    CONST robtarget Target_LetFron3_660:=[[-82.267,-107.387,45.753],[0.430645927,0.216920311,0.57802214,0.658316087],[0,0,0,0],[9E+09,9E+09,9E+09,9E+09,9E+09,9E+09]];
    CONST robtarget Target_LetFron3_670:=[[-81.504,-107.822,44.831],[0.430645927,0.216920311,0.57802214,0.658316087],[0,0,0,0],[9E+09,9E+09,9E+09,9E+09,9E+09,9E+09]];
    CONST robtarget Target_LetFron3_680:=[[-81.6,-107.767,55.109],[0.430645927,0.216920311,0.57802214,0.658316087],[0,0,0,0],[9E+09,9E+09,9E+09,9E+09,9E+09,9E+09]];
    CONST robtarget Target_LetFron3_690:=[[-91.637,-127.746,55.109],[0.430645927,0.216920311,0.57802214,0.658316087],[0,0,0,0],[9E+09,9E+09,9E+09,9E+09,9E+09,9E+09]];
    CONST robtarget Target_LetFron3_700:=[[-88.514,-129.459,54.672],[0.430645927,0.216920311,0.57802214,0.658316087],[0,0,0,0],[9E+09,9E+09,9E+09,9E+09,9E+09,9E+09]];
    CONST robtarget Target_LetFron3_710:=[[-78.514,-109.459,54.672],[0.430645927,0.216920311,0.57802214,0.658316087],[0,0,0,0],[9E+09,9E+09,9E+09,9E+09,9E+09,9E+09]];
    CONST robtarget Target_LetFron3_720:=[[-77.118,-110.187,55.177],[0.430645927,0.216920311,0.57802214,0.658316087],[0,0,0,0],[9E+09,9E+09,9E+09,9E+09,9E+09,9E+09]];
    CONST robtarget Target_LetFron3_730:=[[-75.152,-111.175,55.401],[0.430645927,0.216920311,0.57802214,0.658316087],[0,0,0,0],[9E+09,9E+09,9E+09,9E+09,9E+09,9E+09]];
    CONST robtarget Target_LetFron3_740:=[[-73.482,-111.981,54.982],[0.430645927,0.216920311,0.57802214,0.658316087],[0,0,0,0],[9E+09,9E+09,9E+09,9E+09,9E+09,9E+09]];
    CONST robtarget Target_LetFron3_750:=[[-72.199,-112.579,54.044],[0.430645927,0.216920311,0.57802214,0.658316087],[0,0,0,0],[9E+09,9E+09,9E+09,9E+09,9E+09,9E+09]];
    CONST robtarget Target_LetFron3_760:=[[-71.586,-112.859,52.943],[0.430645927,0.216920311,0.57802214,0.658316087],[0,0,0,0],[9E+09,9E+09,9E+09,9E+09,9E+09,9E+09]];
    CONST robtarget Target_LetFron3_770:=[[-71.209,-113.029,51.815],[0.430645927,0.216920311,0.57802214,0.658316087],[0,0,0,0],[9E+09,9E+09,9E+09,9E+09,9E+09,9E+09]];
    CONST robtarget Target_LetFron3_780:=[[-71.14,-113.06,50.668],[0.430645927,0.216920311,0.57802214,0.658316087],[0,0,0,0],[9E+09,9E+09,9E+09,9E+09,9E+09,9E+09]];
    CONST robtarget Target_LetFron3_790:=[[-71.14,-113.06,49.432],[0.430645927,0.216920311,0.57802214,0.658316087],[0,0,0,0],[9E+09,9E+09,9E+09,9E+09,9E+09,9E+09]];
    CONST robtarget Target_LetFron3_800:=[[-71.288,-112.994,48.254],[0.430645927,0.216920311,0.57802214,0.658316087],[0,0,0,0],[9E+09,9E+09,9E+09,9E+09,9E+09,9E+09]];
    CONST robtarget Target_LetFron3_810:=[[-71.728,-112.794,47.133],[0.430645927,0.216920311,0.57802214,0.658316087],[0,0,0,0],[9E+09,9E+09,9E+09,9E+09,9E+09,9E+09]];
    CONST robtarget Target_LetFron3_820:=[[-72.376,-112.498,46.001],[0.430645927,0.216920311,0.57802214,0.658316087],[0,0,0,0],[9E+09,9E+09,9E+09,9E+09,9E+09,9E+09]];
    CONST robtarget Target_LetFron3_830:=[[-73.318,-112.058,45.279],[0.430645927,0.216920311,0.57802214,0.658316087],[0,0,0,0],[9E+09,9E+09,9E+09,9E+09,9E+09,9E+09]];
    CONST robtarget Target_LetFron3_840:=[[-74.681,-111.405,44.719],[0.430645927,0.216920311,0.57802214,0.658316087],[0,0,0,0],[9E+09,9E+09,9E+09,9E+09,9E+09,9E+09]];
    CONST robtarget Target_LetFron3_850:=[[-75.902,-110.803,44.719],[0.430645927,0.216920311,0.57802214,0.658316087],[0,0,0,0],[9E+09,9E+09,9E+09,9E+09,9E+09,9E+09]];
    CONST robtarget Target_LetFron3_860:=[[-77.054,-110.22,45.141],[0.430645927,0.216920311,0.57802214,0.658316087],[0,0,0,0],[9E+09,9E+09,9E+09,9E+09,9E+09,9E+09]];
    CONST robtarget Target_LetFron3_870:=[[-77.919,-109.772,46.005],[0.430645927,0.216920311,0.57802214,0.658316087],[0,0,0,0],[9E+09,9E+09,9E+09,9E+09,9E+09,9E+09]];
    CONST robtarget Target_LetFron3_880:=[[-78.398,-109.52,46.991],[0.430645927,0.216920311,0.57802214,0.658316087],[0,0,0,0],[9E+09,9E+09,9E+09,9E+09,9E+09,9E+09]];
    CONST robtarget Target_LetFron3_890:=[[-78.609,-109.408,48.208],[0.430645927,0.216920311,0.57802214,0.658316087],[0,0,0,0],[9E+09,9E+09,9E+09,9E+09,9E+09,9E+09]];
    CONST robtarget Target_LetFron3_900:=[[-78.594,-109.416,49.608],[0.430645927,0.216920311,0.57802214,0.658316087],[0,0,0,0],[9E+09,9E+09,9E+09,9E+09,9E+09,9E+09]];
    CONST robtarget Target_LetFron3_910:=[[-78.574,-109.427,49.862],[0.430645927,0.216920311,0.57802214,0.658316087],[0,0,0,0],[9E+09,9E+09,9E+09,9E+09,9E+09,9E+09]];
    CONST robtarget Target_LetFron3_920:=[[-77.106,-110.19,49.869],[0.430645927,0.216920311,0.57802214,0.658316087],[0,0,0,0],[9E+09,9E+09,9E+09,9E+09,9E+09,9E+09]];
    CONST robtarget Target_LetFron3_930:=[[-72.898,-112.255,49.869],[0.430645927,0.216920311,0.57802214,0.658316087],[0,0,0,0],[9E+09,9E+09,9E+09,9E+09,9E+09,9E+09]];
    CONST robtarget Target_LetFron3_940:=[[-82.898,-132.255,49.869],[0.430645927,0.216920311,0.57802214,0.658316087],[0,0,0,0],[9E+09,9E+09,9E+09,9E+09,9E+09,9E+09]];
    CONST robtarget Target_LetFron3_950:=[[-80.313,-133.427,54.778],[0.430645927,0.216920311,0.57802214,0.658316087],[0,0,0,0],[9E+09,9E+09,9E+09,9E+09,9E+09,9E+09]];
    CONST robtarget Target_LetFron3_960:=[[-70.313,-113.427,54.778],[0.430645927,0.216920311,0.57802214,0.658316087],[0,0,0,0],[9E+09,9E+09,9E+09,9E+09,9E+09,9E+09]];
    CONST robtarget Target_LetFron3_970:=[[-68.992,-113.999,55.279],[0.430645927,0.216920311,0.57802214,0.658316087],[0,0,0,0],[9E+09,9E+09,9E+09,9E+09,9E+09,9E+09]];
    CONST robtarget Target_LetFron3_980:=[[-67.664,-114.556,55.401],[0.430645927,0.216920311,0.57802214,0.658316087],[0,0,0,0],[9E+09,9E+09,9E+09,9E+09,9E+09,9E+09]];
    CONST robtarget Target_LetFron3_990:=[[-66.498,-115.03,55.08],[0.430645927,0.216920311,0.57802214,0.658316087],[0,0,0,0],[9E+09,9E+09,9E+09,9E+09,9E+09,9E+09]];
    CONST robtarget Target_LetFron3_1000:=[[-65.468,-115.437,54.06],[0.430645927,0.216920311,0.57802214,0.658316087],[0,0,0,0],[9E+09,9E+09,9E+09,9E+09,9E+09,9E+09]];
    CONST robtarget Target_LetFron3_1010:=[[-65.245,-115.524,53.314],[0.430645927,0.216920311,0.57802214,0.658316087],[0,0,0,0],[9E+09,9E+09,9E+09,9E+09,9E+09,9E+09]];
    CONST robtarget Target_LetFron3_1020:=[[-65.368,-115.476,43.276],[0.430645927,0.216920311,0.57802214,0.658316087],[0,0,0,0],[9E+09,9E+09,9E+09,9E+09,9E+09,9E+09]];
    CONST robtarget Target_LetFron3_1030:=[[-65.313,-115.498,44.991],[0.430645927,0.216920311,0.57802214,0.658316087],[0,0,0,0],[9E+09,9E+09,9E+09,9E+09,9E+09,9E+09]];
    CONST robtarget Target_LetFron3_1040:=[[-63.93,-116.026,45.188],[0.430645927,0.216920311,0.57802214,0.658316087],[0,0,0,0],[9E+09,9E+09,9E+09,9E+09,9E+09,9E+09]];
    CONST robtarget Target_LetFron3_1050:=[[-70.13,-113.508,44.989],[0.430645927,0.216920311,0.57802214,0.658316087],[0,0,0,0],[9E+09,9E+09,9E+09,9E+09,9E+09,9E+09]];
    CONST robtarget Target_LetFron3_1060:=[[-80.13,-133.508,44.989],[0.430645927,0.216920311,0.57802214,0.658316087],[0,0,0,0],[9E+09,9E+09,9E+09,9E+09,9E+09,9E+09]];
    CONST robtarget Target_LetFron3_1070:=[[-72.339,-136.611,45.952],[0.430645927,0.216920311,0.57802214,0.658316087],[0,0,0,0],[9E+09,9E+09,9E+09,9E+09,9E+09,9E+09]];
    CONST robtarget Target_LetFron3_1080:=[[-62.36,-116.604,45.863],[0.430645927,0.216920311,0.57802214,0.658316087],[0,0,0,0],[9E+09,9E+09,9E+09,9E+09,9E+09,9E+09]];
    CONST robtarget Target_LetFron3_1090:=[[-60.366,-117.303,44.736],[0.430645927,0.216920311,0.57802214,0.658316087],[0,0,0,0],[9E+09,9E+09,9E+09,9E+09,9E+09,9E+09]];
    CONST robtarget Target_LetFron3_1100:=[[-58.61,-117.888,44.82],[0.430645927,0.216920311,0.57802214,0.658316087],[0,0,0,0],[9E+09,9E+09,9E+09,9E+09,9E+09,9E+09]];
    CONST robtarget Target_LetFron3_1110:=[[-56.667,-118.501,45.956],[0.430645927,0.216920311,0.57802214,0.658316087],[0,0,0,0],[9E+09,9E+09,9E+09,9E+09,9E+09,9E+09]];
    CONST robtarget Target_LetFron3_1120:=[[-56.029,-118.695,47.133],[0.430645927,0.216920311,0.57802214,0.658316087],[0,0,0,0],[9E+09,9E+09,9E+09,9E+09,9E+09,9E+09]];
    CONST robtarget Target_LetFron3_1130:=[[-56.121,-118.667,48.621],[0.430645927,0.216920311,0.57802214,0.658316087],[0,0,0,0],[9E+09,9E+09,9E+09,9E+09,9E+09,9E+09]];
    CONST robtarget Target_LetFron3_1140:=[[-56.545,-118.539,49.359],[0.430645927,0.216920311,0.57802214,0.658316087],[0,0,0,0],[9E+09,9E+09,9E+09,9E+09,9E+09,9E+09]];
    CONST robtarget Target_LetFron3_1150:=[[-57.437,-118.262,50.034],[0.430645927,0.216920311,0.57802214,0.658316087],[0,0,0,0],[9E+09,9E+09,9E+09,9E+09,9E+09,9E+09]];
    CONST robtarget Target_LetFron3_1160:=[[-58.505,-117.922,50.535],[0.430645927,0.216920311,0.57802214,0.658316087],[0,0,0,0],[9E+09,9E+09,9E+09,9E+09,9E+09,9E+09]];
    CONST robtarget Target_LetFron3_1170:=[[-59.869,-117.471,51.117],[0.430645927,0.216920311,0.57802214,0.658316087],[0,0,0,0],[9E+09,9E+09,9E+09,9E+09,9E+09,9E+09]];
    CONST robtarget Target_LetFron3_1180:=[[-60.318,-117.319,51.376],[0.430645927,0.216920311,0.57802214,0.658316087],[0,0,0,0],[9E+09,9E+09,9E+09,9E+09,9E+09,9E+09]];
    CONST robtarget Target_LetFron3_1190:=[[-62.669,-116.492,52.048],[0.430645927,0.216920311,0.57802214,0.658316087],[0,0,0,0],[9E+09,9E+09,9E+09,9E+09,9E+09,9E+09]];
    CONST robtarget Target_LetFron3_1200:=[[-62.602,-116.516,52.834],[0.430645927,0.216920311,0.57802214,0.658316087],[0,0,0,0],[9E+09,9E+09,9E+09,9E+09,9E+09,9E+09]];
    CONST robtarget Target_LetFron3_1210:=[[-62.228,-116.651,53.814],[0.430645927,0.216920311,0.57802214,0.658316087],[0,0,0,0],[9E+09,9E+09,9E+09,9E+09,9E+09,9E+09]];
    CONST robtarget Target_LetFron3_1220:=[[-61.449,-116.928,54.619],[0.430645927,0.216920311,0.57802214,0.658316087],[0,0,0,0],[9E+09,9E+09,9E+09,9E+09,9E+09,9E+09]];
    CONST robtarget Target_LetFron3_1230:=[[-60.216,-117.353,55.205],[0.430645927,0.216920311,0.57802214,0.658316087],[0,0,0,0],[9E+09,9E+09,9E+09,9E+09,9E+09,9E+09]];
    CONST robtarget Target_LetFron3_1240:=[[-58.271,-117.997,55.4],[0.430645927,0.216920311,0.57802214,0.658316087],[0,0,0,0],[9E+09,9E+09,9E+09,9E+09,9E+09,9E+09]];
    CONST robtarget Target_LetFron3_1250:=[[-56.602,-118.521,55.079],[0.430645927,0.216920311,0.57802214,0.658316087],[0,0,0,0],[9E+09,9E+09,9E+09,9E+09,9E+09,9E+09]];
    CONST robtarget Target_LetFron3_1260:=[[-55.798,-118.764,54.785],[0.430645927,0.216920311,0.57802214,0.658316087],[0,0,0,0],[9E+09,9E+09,9E+09,9E+09,9E+09,9E+09]];
    CONST robtarget Target_LetFron3_1270:=[[-65.797,-138.765,54.792],[0.430645927,0.216920311,0.57802214,0.658316087],[0,0,0,0],[9E+09,9E+09,9E+09,9E+09,9E+09,9E+09]];
    CONST robtarget Target_LetFron3_1280:=[[-62.847,-139.607,55.109],[0.430645927,0.216920311,0.57802214,0.658316087],[0,0,0,0],[9E+09,9E+09,9E+09,9E+09,9E+09,9E+09]];
    CONST robtarget Target_LetFron3_1290:=[[-52.847,-119.607,55.109],[0.430645927,0.216920311,0.57802214,0.658316087],[0,0,0,0],[9E+09,9E+09,9E+09,9E+09,9E+09,9E+09]];
    CONST robtarget Target_LetFron3_1300:=[[-52.608,-119.672,44.874],[0.430645927,0.216920311,0.57802214,0.658316087],[0,0,0,0],[9E+09,9E+09,9E+09,9E+09,9E+09,9E+09]];
    CONST robtarget Target_LetFron3_1310:=[[-62.608,-139.672,44.874],[0.430645927,0.216920311,0.57802214,0.658316087],[0,0,0,0],[9E+09,9E+09,9E+09,9E+09,9E+09,9E+09]];
    CONST robtarget Target_LetFron3_1320:=[[-62.417,-139.723,40.356],[0.430645927,0.216920311,0.57802214,0.658316087],[0,0,0,0],[9E+09,9E+09,9E+09,9E+09,9E+09,9E+09]];
    CONST robtarget Target_LetFron3_1330:=[[-52.574,-119.681,40.311],[0.430645927,0.216920311,0.57802214,0.658316087],[0,0,0,0],[9E+09,9E+09,9E+09,9E+09,9E+09,9E+09]];
    CONST robtarget Target_LetFron3_1340:=[[-62.574,-139.681,40.311],[0.430645927,0.216920311,0.57802214,0.658316087],[0,0,0,0],[9E+09,9E+09,9E+09,9E+09,9E+09,9E+09]];
    CONST robtarget Target_LetFron3_1350:=[[-58.595,-140.685,42.493],[0.430645927,0.216920311,0.57802214,0.658316087],[0,0,0,0],[9E+09,9E+09,9E+09,9E+09,9E+09,9E+09]];
    CONST robtarget Target_LetFron3_1360:=[[-48.595,-120.685,42.493],[0.430645927,0.216920311,0.57802214,0.658316087],[0,0,0,0],[9E+09,9E+09,9E+09,9E+09,9E+09,9E+09]];
    CONST robtarget Target_LetFron3_1370:=[[-42.535,-121.952,41.813],[0.430645927,0.216920311,0.57802214,0.658316087],[0,0,0,0],[9E+09,9E+09,9E+09,9E+09,9E+09,9E+09]];
    CONST robtarget Target_LetFron3_1380:=[[-41.416,-122.152,42.942],[0.430645927,0.216920311,0.57802214,0.658316087],[0,0,0,0],[9E+09,9E+09,9E+09,9E+09,9E+09,9E+09]];
    CONST robtarget Target_LetFron3_1390:=[[-40.861,-122.247,44.157],[0.430645927,0.216920311,0.57802214,0.658316087],[0,0,0,0],[9E+09,9E+09,9E+09,9E+09,9E+09,9E+09]];
    CONST robtarget Target_LetFron3_1400:=[[-40.861,-122.247,45.481],[0.430645927,0.216920311,0.57802214,0.658316087],[0,0,0,0],[9E+09,9E+09,9E+09,9E+09,9E+09,9E+09]];
    CONST robtarget Target_LetFron3_1410:=[[-41.204,-122.188,46.641],[0.430645927,0.216920311,0.57802214,0.658316087],[0,0,0,0],[9E+09,9E+09,9E+09,9E+09,9E+09,9E+09]];
    CONST robtarget Target_LetFron3_1420:=[[-41.998,-122.049,47.583],[0.430645927,0.216920311,0.57802214,0.658316087],[0,0,0,0],[9E+09,9E+09,9E+09,9E+09,9E+09,9E+09]];
    CONST robtarget Target_LetFron3_1430:=[[-43.35,-121.797,48.403],[0.430645927,0.216920311,0.57802214,0.658316087],[0,0,0,0],[9E+09,9E+09,9E+09,9E+09,9E+09,9E+09]];
    CONST robtarget Target_LetFron3_1440:=[[-44.844,-121.506,49.112],[0.430645927,0.216920311,0.57802214,0.658316087],[0,0,0,0],[9E+09,9E+09,9E+09,9E+09,9E+09,9E+09]];
    CONST robtarget Target_LetFron3_1450:=[[-46.229,-121.217,49.939],[0.430645927,0.216920311,0.57802214,0.658316087],[0,0,0,0],[9E+09,9E+09,9E+09,9E+09,9E+09,9E+09]];
    CONST robtarget Target_LetFron3_1460:=[[-49.035,-120.581,50.611],[0.430645927,0.216920311,0.57802214,0.658316087],[0,0,0,0],[9E+09,9E+09,9E+09,9E+09,9E+09,9E+09]];
    CONST robtarget Target_LetFron3_1470:=[[-48.955,-120.6,52.318],[0.430645927,0.216920311,0.57802214,0.658316087],[0,0,0,0],[9E+09,9E+09,9E+09,9E+09,9E+09,9E+09]];
    CONST robtarget Target_LetFron3_1480:=[[-48.452,-120.719,53.355],[0.430645927,0.216920311,0.57802214,0.658316087],[0,0,0,0],[9E+09,9E+09,9E+09,9E+09,9E+09,9E+09]];
    CONST robtarget Target_LetFron3_1490:=[[-47.435,-120.951,54.415],[0.430645927,0.216920311,0.57802214,0.658316087],[0,0,0,0],[9E+09,9E+09,9E+09,9E+09,9E+09,9E+09]];
    CONST robtarget Target_LetFron3_1500:=[[-45.861,-121.294,55.128],[0.430645927,0.216920311,0.57802214,0.658316087],[0,0,0,0],[9E+09,9E+09,9E+09,9E+09,9E+09,9E+09]];
    CONST robtarget Target_LetFron3_1510:=[[-43.532,-121.765,55.401],[0.430645927,0.216920311,0.57802214,0.658316087],[0,0,0,0],[9E+09,9E+09,9E+09,9E+09,9E+09,9E+09]];
    CONST robtarget Target_LetFron3_1520:=[[-41.726,-122.098,55.154],[0.430645927,0.216920311,0.57802214,0.658316087],[0,0,0,0],[9E+09,9E+09,9E+09,9E+09,9E+09,9E+09]];
    CONST robtarget Target_LetFron3_1530:=[[-40.575,-122.295,54.72],[0.430645927,0.216920311,0.57802214,0.658316087],[0,0,0,0],[9E+09,9E+09,9E+09,9E+09,9E+09,9E+09]];
    CONST robtarget Target_LetFron3_1540:=[[-50.576,-142.295,54.717],[0.430645927,0.216920311,0.57802214,0.658316087],[0,0,0,0],[9E+09,9E+09,9E+09,9E+09,9E+09,9E+09]];
    CONST robtarget Target_LetFron3_1550:=[[-43.98,-143.216,54.592],[0.430645927,0.216920311,0.57802214,0.658316087],[0,0,0,0],[9E+09,9E+09,9E+09,9E+09,9E+09,9E+09]];
    CONST robtarget Target_LetFron3_1560:=[[-33.98,-123.216,54.592],[0.430645927,0.216920311,0.57802214,0.658316087],[0,0,0,0],[9E+09,9E+09,9E+09,9E+09,9E+09,9E+09]];
    CONST robtarget Target_LetFron3_1570:=[[-32.448,-123.378,55.116],[0.430645927,0.216920311,0.57802214,0.658316087],[0,0,0,0],[9E+09,9E+09,9E+09,9E+09,9E+09,9E+09]];
    CONST robtarget Target_LetFron3_1580:=[[-30.55,-123.554,55.401],[0.430645927,0.216920311,0.57802214,0.658316087],[0,0,0,0],[9E+09,9E+09,9E+09,9E+09,9E+09,9E+09]];
    CONST robtarget Target_LetFron3_1590:=[[-28.936,-123.68,55.282],[0.430645927,0.216920311,0.57802214,0.658316087],[0,0,0,0],[9E+09,9E+09,9E+09,9E+09,9E+09,9E+09]];
    CONST robtarget Target_LetFron3_1600:=[[-27.719,-123.761,54.742],[0.430645927,0.216920311,0.57802214,0.658316087],[0,0,0,0],[9E+09,9E+09,9E+09,9E+09,9E+09,9E+09]];
    CONST robtarget Target_LetFron3_1610:=[[-26.596,-123.826,53.8],[0.430645927,0.216920311,0.57802214,0.658316087],[0,0,0,0],[9E+09,9E+09,9E+09,9E+09,9E+09,9E+09]];
    CONST robtarget Target_LetFron3_1620:=[[-25.968,-123.857,52.688],[0.430645927,0.216920311,0.57802214,0.658316087],[0,0,0,0],[9E+09,9E+09,9E+09,9E+09,9E+09,9E+09]];
    CONST robtarget Target_LetFron3_1630:=[[-25.618,-123.874,50.949],[0.430645927,0.216920311,0.57802214,0.658316087],[0,0,0,0],[9E+09,9E+09,9E+09,9E+09,9E+09,9E+09]];
    CONST robtarget Target_LetFron3_1640:=[[-25.618,-123.874,49.368],[0.430645927,0.216920311,0.57802214,0.658316087],[0,0,0,0],[9E+09,9E+09,9E+09,9E+09,9E+09,9E+09]];
    CONST robtarget Target_LetFron3_1650:=[[-25.967,-123.858,47.76],[0.430645927,0.216920311,0.57802214,0.658316087],[0,0,0,0],[9E+09,9E+09,9E+09,9E+09,9E+09,9E+09]];
    CONST robtarget Target_LetFron3_1660:=[[-26.976,-123.805,46.001],[0.430645927,0.216920311,0.57802214,0.658316087],[0,0,0,0],[9E+09,9E+09,9E+09,9E+09,9E+09,9E+09]];
    CONST robtarget Target_LetFron3_1670:=[[-28.333,-123.722,45.081],[0.430645927,0.216920311,0.57802214,0.658316087],[0,0,0,0],[9E+09,9E+09,9E+09,9E+09,9E+09,9E+09]];
    CONST robtarget Target_LetFron3_1680:=[[-29.666,-123.626,44.719],[0.430645927,0.216920311,0.57802214,0.658316087],[0,0,0,0],[9E+09,9E+09,9E+09,9E+09,9E+09,9E+09]];
    CONST robtarget Target_LetFron3_1690:=[[-30.876,-123.526,44.719],[0.430645927,0.216920311,0.57802214,0.658316087],[0,0,0,0],[9E+09,9E+09,9E+09,9E+09,9E+09,9E+09]];
    CONST robtarget Target_LetFron3_1700:=[[-32.317,-123.392,45.206],[0.430645927,0.216920311,0.57802214,0.658316087],[0,0,0,0],[9E+09,9E+09,9E+09,9E+09,9E+09,9E+09]];
    CONST robtarget Target_LetFron3_1710:=[[-32.996,-123.323,45.821],[0.430645927,0.216920311,0.57802214,0.658316087],[0,0,0,0],[9E+09,9E+09,9E+09,9E+09,9E+09,9E+09]];
    CONST robtarget Target_LetFron3_1720:=[[-33.54,-123.265,46.556],[0.430645927,0.216920311,0.57802214,0.658316087],[0,0,0,0],[9E+09,9E+09,9E+09,9E+09,9E+09,9E+09]];
    CONST robtarget Target_LetFron3_1730:=[[-33.887,-123.226,47.949],[0.430645927,0.216920311,0.57802214,0.658316087],[0,0,0,0],[9E+09,9E+09,9E+09,9E+09,9E+09,9E+09]];
    CONST robtarget Target_LetFron3_1740:=[[-33.912,-123.223,49.284],[0.430645927,0.216920311,0.57802214,0.658316087],[0,0,0,0],[9E+09,9E+09,9E+09,9E+09,9E+09,9E+09]];
    CONST robtarget Target_LetFron3_1750:=[[-33.868,-123.228,49.869],[0.430645927,0.216920311,0.57802214,0.658316087],[0,0,0,0],[9E+09,9E+09,9E+09,9E+09,9E+09,9E+09]];
    CONST robtarget Target_LetFron3_1760:=[[-27.55,-123.772,49.869],[0.430645927,0.216920311,0.57802214,0.658316087],[0,0,0,0],[9E+09,9E+09,9E+09,9E+09,9E+09,9E+09]];
    CONST robtarget Target_LetFron3_1770:=[[-37.55,-143.772,49.897],[0.430645927,0.216920311,0.57802214,0.658316087],[0,0,0,0],[9E+09,9E+09,9E+09,9E+09,9E+09,9E+09]];
    CONST robtarget Target_LetFron3_1780:=[[-31.259,-143.994,45.099],[0.430645927,0.216920311,0.57802214,0.658316087],[0,0,0,0],[9E+09,9E+09,9E+09,9E+09,9E+09,9E+09]];
    CONST robtarget Target_LetFron3_1790:=[[-21.259,-123.994,45.14],[0.430645927,0.216920311,0.57802214,0.658316087],[0,0,0,0],[9E+09,9E+09,9E+09,9E+09,9E+09,9E+09]];
    CONST robtarget Target_LetFron3_1800:=[[-19.408,-123.999,44.719],[0.430645927,0.216920311,0.57802214,0.658316087],[0,0,0,0],[9E+09,9E+09,9E+09,9E+09,9E+09,9E+09]];
    CONST robtarget Target_LetFron3_1810:=[[-17.893,-123.982,44.831],[0.430645927,0.216920311,0.57802214,0.658316087],[0,0,0,0],[9E+09,9E+09,9E+09,9E+09,9E+09,9E+09]];
    CONST robtarget Target_LetFron3_1820:=[[-16.252,-123.944,45.604],[0.430645927,0.216920311,0.57802214,0.658316087],[0,0,0,0],[9E+09,9E+09,9E+09,9E+09,9E+09,9E+09]];
    CONST robtarget Target_LetFron3_1830:=[[-15.038,-123.901,46.903],[0.430645927,0.216920311,0.57802214,0.658316087],[0,0,0,0],[9E+09,9E+09,9E+09,9E+09,9E+09,9E+09]];
    CONST robtarget Target_LetFron3_1840:=[[-14.306,-123.87,48.941],[0.430645927,0.216920311,0.57802214,0.658316087],[0,0,0,0],[9E+09,9E+09,9E+09,9E+09,9E+09,9E+09]];
    CONST robtarget Target_LetFron3_1850:=[[-14.248,-123.868,50.838],[0.430645927,0.216920311,0.57802214,0.658316087],[0,0,0,0],[9E+09,9E+09,9E+09,9E+09,9E+09,9E+09]];
    CONST robtarget Target_LetFron3_1860:=[[-14.656,-123.886,52.859],[0.430645927,0.216920311,0.57802214,0.658316087],[0,0,0,0],[9E+09,9E+09,9E+09,9E+09,9E+09,9E+09]];
    CONST robtarget Target_LetFron3_1870:=[[-15.358,-123.914,54.174],[0.430645927,0.216920311,0.57802214,0.658316087],[0,0,0,0],[9E+09,9E+09,9E+09,9E+09,9E+09,9E+09]];
    CONST robtarget Target_LetFron3_1880:=[[-16.312,-123.946,54.884],[0.430645927,0.216920311,0.57802214,0.658316087],[0,0,0,0],[9E+09,9E+09,9E+09,9E+09,9E+09,9E+09]];
    CONST robtarget Target_LetFron3_1890:=[[-17.794,-123.981,55.401],[0.430645927,0.216920311,0.57802214,0.658316087],[0,0,0,0],[9E+09,9E+09,9E+09,9E+09,9E+09,9E+09]];
    CONST robtarget Target_LetFron3_1900:=[[-18.988,-123.996,55.337],[0.430645927,0.216920311,0.57802214,0.658316087],[0,0,0,0],[9E+09,9E+09,9E+09,9E+09,9E+09,9E+09]];
    CONST robtarget Target_LetFron3_1910:=[[-20.839,-123.997,54.644],[0.430645927,0.216920311,0.57802214,0.658316087],[0,0,0,0],[9E+09,9E+09,9E+09,9E+09,9E+09,9E+09]];
    CONST robtarget Target_LetFron3_1920:=[[-21.239,-123.994,54.414],[0.430645927,0.216920311,0.57802214,0.658316087],[0,0,0,0],[9E+09,9E+09,9E+09,9E+09,9E+09,9E+09]];
    CONST robtarget Target_LetFron3_1930:=[[-22.525,-123.974,55.243],[0.430645927,0.216920311,0.57802214,0.658316087],[0,0,0,0],[9E+09,9E+09,9E+09,9E+09,9E+09,9E+09]];
    CONST robtarget Target_LetFron3_1940:=[[-22.191,-123.98,39.777],[0.430645927,0.216920311,0.57802214,0.658316087],[0,0,0,0],[9E+09,9E+09,9E+09,9E+09,9E+09,9E+09]];
    CONST robtarget Target_LetFron3_1950:=[[-32.321,-143.978,39.756],[0.430645927,0.216920311,0.57802214,0.658316087],[0,0,0,0],[9E+09,9E+09,9E+09,9E+09,9E+09,9E+09]];
    CONST robtarget Target_LetFron3_1960:=[[-12.321,-144.978,-58.244],[0.443836724,0.190106418,0.616719914,0.621711396],[0,0,0,0],[9E+09,9E+09,9E+09,9E+09,9E+09,9E+09]];
    !***********************************************************
    !Dibujo cuarto cuadrante de letrero frontal
    CONST robtarget Target_LetFron4_10:=[[-8.95,-145.995,82.097],[0.503297686,0.226891536,0.589713525,0.58944858],[0,0,0,0],[9E+09,9E+09,9E+09,9E+09,9E+09,9E+09]];
    CONST robtarget Target_LetFron4_20:=[[-18.95,-125.995,82.097],[0.503297686,0.226891536,0.589713525,0.58944858],[0,0,0,0],[9E+09,9E+09,9E+09,9E+09,9E+09,9E+09]];
    CONST robtarget Target_LetFron4_30:=[[-19.003,-125.994,68.333],[0.503297686,0.226891536,0.589713525,0.58944858],[0,0,0,0],[9E+09,9E+09,9E+09,9E+09,9E+09,9E+09]];
    CONST robtarget Target_LetFron4_40:=[[-23.592,-125.948,68.333],[0.503297686,0.226891536,0.589713525,0.58944858],[0,0,0,0],[9E+09,9E+09,9E+09,9E+09,9E+09,9E+09]];
    CONST robtarget Target_LetFron4_50:=[[-25.245,-125.89,69.103],[0.503297686,0.226891536,0.589713525,0.58944858],[0,0,0,0],[9E+09,9E+09,9E+09,9E+09,9E+09,9E+09]];
    CONST robtarget Target_LetFron4_60:=[[-26.403,-125.836,70.475],[0.503297686,0.226891536,0.589713525,0.58944858],[0,0,0,0],[9E+09,9E+09,9E+09,9E+09,9E+09,9E+09]];
    CONST robtarget Target_LetFron4_70:=[[-26.7,-125.82,71.985],[0.503297686,0.226891536,0.589713525,0.58944858],[0,0,0,0],[9E+09,9E+09,9E+09,9E+09,9E+09,9E+09]];
    CONST robtarget Target_LetFron4_80:=[[-26.314,-125.84,73.908],[0.503297686,0.226891536,0.589713525,0.58944858],[0,0,0,0],[9E+09,9E+09,9E+09,9E+09,9E+09,9E+09]];
    CONST robtarget Target_LetFron4_90:=[[-24.963,-125.901,75.447],[0.503297686,0.226891536,0.589713525,0.58944858],[0,0,0,0],[9E+09,9E+09,9E+09,9E+09,9E+09,9E+09]];
    CONST robtarget Target_LetFron4_100:=[[-21.051,-125.996,76.407],[0.503297686,0.226891536,0.589713525,0.58944858],[0,0,0,0],[9E+09,9E+09,9E+09,9E+09,9E+09,9E+09]];
    CONST robtarget Target_LetFron4_110:=[[-22.431,-125.976,76.317],[0.503297686,0.226891536,0.589713525,0.58944858],[0,0,0,0],[9E+09,9E+09,9E+09,9E+09,9E+09,9E+09]];
    CONST robtarget Target_LetFron4_120:=[[-26.29,-125.841,82.097],[0.503297686,0.226891536,0.589713525,0.58944858],[0,0,0,0],[9E+09,9E+09,9E+09,9E+09,9E+09,9E+09]];
    CONST robtarget Target_LetFron4_130:=[[-36.29,-145.841,82.097],[0.503297686,0.226891536,0.589713525,0.58944858],[0,0,0,0],[9E+09,9E+09,9E+09,9E+09,9E+09,9E+09]];
    CONST robtarget Target_LetFron4_140:=[[-42.667,-145.355,82.283],[0.503297686,0.226891536,0.589713525,0.58944858],[0,0,0,0],[9E+09,9E+09,9E+09,9E+09,9E+09,9E+09]];
    CONST robtarget Target_LetFron4_150:=[[-32.667,-125.355,82.283],[0.503297686,0.226891536,0.589713525,0.58944858],[0,0,0,0],[9E+09,9E+09,9E+09,9E+09,9E+09,9E+09]];
    CONST robtarget Target_LetFron4_160:=[[-34.857,-125.114,82.316],[0.503297686,0.226891536,0.589713525,0.58944858],[0,0,0,0],[9E+09,9E+09,9E+09,9E+09,9E+09,9E+09]];
    CONST robtarget Target_LetFron4_170:=[[-36.701,-124.879,81.437],[0.503297686,0.226891536,0.589713525,0.58944858],[0,0,0,0],[9E+09,9E+09,9E+09,9E+09,9E+09,9E+09]];
    CONST robtarget Target_LetFron4_180:=[[-37.577,-124.758,80.559],[0.503297686,0.226891536,0.589713525,0.58944858],[0,0,0,0],[9E+09,9E+09,9E+09,9E+09,9E+09,9E+09]];
    CONST robtarget Target_LetFron4_190:=[[-38.397,-124.639,78.755],[0.503297686,0.226891536,0.589713525,0.58944858],[0,0,0,0],[9E+09,9E+09,9E+09,9E+09,9E+09,9E+09]];
    CONST robtarget Target_LetFron4_200:=[[-38.556,-124.615,76.834],[0.503297686,0.226891536,0.589713525,0.58944858],[0,0,0,0],[9E+09,9E+09,9E+09,9E+09,9E+09,9E+09]];
    CONST robtarget Target_LetFron4_210:=[[-38.535,-124.618,75.633],[0.503297686,0.226891536,0.589713525,0.58944858],[0,0,0,0],[9E+09,9E+09,9E+09,9E+09,9E+09,9E+09]];
    CONST robtarget Target_LetFron4_220:=[[-38.089,-124.684,74.246],[0.503297686,0.226891536,0.589713525,0.58944858],[0,0,0,0],[9E+09,9E+09,9E+09,9E+09,9E+09,9E+09]];
    CONST robtarget Target_LetFron4_230:=[[-37.456,-124.775,73.108],[0.503297686,0.226891536,0.589713525,0.58944858],[0,0,0,0],[9E+09,9E+09,9E+09,9E+09,9E+09,9E+09]];
    CONST robtarget Target_LetFron4_240:=[[-36.441,-124.914,72.314],[0.503297686,0.226891536,0.589713525,0.58944858],[0,0,0,0],[9E+09,9E+09,9E+09,9E+09,9E+09,9E+09]];
    CONST robtarget Target_LetFron4_250:=[[-35.37,-125.051,71.858],[0.503297686,0.226891536,0.589713525,0.58944858],[0,0,0,0],[9E+09,9E+09,9E+09,9E+09,9E+09,9E+09]];
    CONST robtarget Target_LetFron4_260:=[[-33.892,-125.226,71.706],[0.503297686,0.226891536,0.589713525,0.58944858],[0,0,0,0],[9E+09,9E+09,9E+09,9E+09,9E+09,9E+09]];
    CONST robtarget Target_LetFron4_270:=[[-32.661,-125.357,71.87],[0.503297686,0.226891536,0.589713525,0.58944858],[0,0,0,0],[9E+09,9E+09,9E+09,9E+09,9E+09,9E+09]];
    CONST robtarget Target_LetFron4_280:=[[-31.413,-125.478,72.359],[0.503297686,0.226891536,0.589713525,0.58944858],[0,0,0,0],[9E+09,9E+09,9E+09,9E+09,9E+09,9E+09]];
    CONST robtarget Target_LetFron4_290:=[[-30.454,-125.562,73.003],[0.503297686,0.226891536,0.589713525,0.58944858],[0,0,0,0],[9E+09,9E+09,9E+09,9E+09,9E+09,9E+09]];
    CONST robtarget Target_LetFron4_300:=[[-29.503,-125.638,74.523],[0.503297686,0.226891536,0.589713525,0.58944858],[0,0,0,0],[9E+09,9E+09,9E+09,9E+09,9E+09,9E+09]];
    CONST robtarget Target_LetFron4_310:=[[-29.14,-125.665,75.942],[0.503297686,0.226891536,0.589713525,0.58944858],[0,0,0,0],[9E+09,9E+09,9E+09,9E+09,9E+09,9E+09]];
    CONST robtarget Target_LetFron4_320:=[[-29.014,-125.675,77.239],[0.503297686,0.226891536,0.589713525,0.58944858],[0,0,0,0],[9E+09,9E+09,9E+09,9E+09,9E+09,9E+09]];
    CONST robtarget Target_LetFron4_330:=[[-29.16,-125.664,78.757],[0.503297686,0.226891536,0.589713525,0.58944858],[0,0,0,0],[9E+09,9E+09,9E+09,9E+09,9E+09,9E+09]];
    CONST robtarget Target_LetFron4_340:=[[-29.598,-125.631,80.028],[0.503297686,0.226891536,0.589713525,0.58944858],[0,0,0,0],[9E+09,9E+09,9E+09,9E+09,9E+09,9E+09]];
    CONST robtarget Target_LetFron4_350:=[[-30.232,-125.58,80.936],[0.503297686,0.226891536,0.589713525,0.58944858],[0,0,0,0],[9E+09,9E+09,9E+09,9E+09,9E+09,9E+09]];
    CONST robtarget Target_LetFron4_360:=[[-31.211,-125.496,81.782],[0.503297686,0.226891536,0.589713525,0.58944858],[0,0,0,0],[9E+09,9E+09,9E+09,9E+09,9E+09,9E+09]];
    CONST robtarget Target_LetFron4_370:=[[-32.734,-125.348,82.291],[0.503297686,0.226891536,0.589713525,0.58944858],[0,0,0,0],[9E+09,9E+09,9E+09,9E+09,9E+09,9E+09]];
    CONST robtarget Target_LetFron4_380:=[[-42.734,-145.348,82.291],[0.503297686,0.226891536,0.589713525,0.58944858],[0,0,0,0],[9E+09,9E+09,9E+09,9E+09,9E+09,9E+09]];
    CONST robtarget Target_LetFron4_390:=[[-53.051,-143.856,72.591],[0.492892784,0.289203693,0.528592352,0.627700607],[0,0,0,0],[9E+09,9E+09,9E+09,9E+09,9E+09,9E+09]];
    CONST robtarget Target_LetFron4_400:=[[-43.051,-123.856,72.591],[0.492892784,0.289203693,0.528592352,0.627700607],[0,0,0,0],[9E+09,9E+09,9E+09,9E+09,9E+09,9E+09]];
    CONST robtarget Target_LetFron4_410:=[[-45.7,-123.329,71.706],[0.492892784,0.289203693,0.528592352,0.627700607],[0,0,0,0],[9E+09,9E+09,9E+09,9E+09,9E+09,9E+09]];
    CONST robtarget Target_LetFron4_420:=[[-46.898,-123.072,71.822],[0.492892784,0.289203693,0.528592352,0.627700607],[0,0,0,0],[9E+09,9E+09,9E+09,9E+09,9E+09,9E+09]];
    CONST robtarget Target_LetFron4_430:=[[-48.129,-122.794,72.468],[0.492892784,0.289203693,0.528592352,0.627700607],[0,0,0,0],[9E+09,9E+09,9E+09,9E+09,9E+09,9E+09]];
    CONST robtarget Target_LetFron4_440:=[[-49.172,-122.548,73.865],[0.492892784,0.289203693,0.528592352,0.627700607],[0,0,0,0],[9E+09,9E+09,9E+09,9E+09,9E+09,9E+09]];
    CONST robtarget Target_LetFron4_450:=[[-49.762,-122.405,76.003],[0.492892784,0.289203693,0.528592352,0.627700607],[0,0,0,0],[9E+09,9E+09,9E+09,9E+09,9E+09,9E+09]];
    CONST robtarget Target_LetFron4_460:=[[-49.705,-122.419,78.093],[0.492892784,0.289203693,0.528592352,0.627700607],[0,0,0,0],[9E+09,9E+09,9E+09,9E+09,9E+09,9E+09]];
    CONST robtarget Target_LetFron4_470:=[[-49.07,-122.573,80.012],[0.492892784,0.289203693,0.528592352,0.627700607],[0,0,0,0],[9E+09,9E+09,9E+09,9E+09,9E+09,9E+09]];
    CONST robtarget Target_LetFron4_480:=[[-47.496,-122.938,81.652],[0.492892784,0.289203693,0.528592352,0.627700607],[0,0,0,0],[9E+09,9E+09,9E+09,9E+09,9E+09,9E+09]];
    CONST robtarget Target_LetFron4_490:=[[-45.602,-123.35,82.389],[0.492892784,0.289203693,0.528592352,0.627700607],[0,0,0,0],[9E+09,9E+09,9E+09,9E+09,9E+09,9E+09]];
    CONST robtarget Target_LetFron4_500:=[[-43.633,-123.746,82.209],[0.492892784,0.289203693,0.528592352,0.627700607],[0,0,0,0],[9E+09,9E+09,9E+09,9E+09,9E+09,9E+09]];
    CONST robtarget Target_LetFron4_510:=[[-42.513,-123.956,81.879],[0.492892784,0.289203693,0.528592352,0.627700607],[0,0,0,0],[9E+09,9E+09,9E+09,9E+09,9E+09,9E+09]];
    CONST robtarget Target_LetFron4_520:=[[-41.582,-124.123,82.545],[0.492892784,0.289203693,0.528592352,0.627700607],[0,0,0,0],[9E+09,9E+09,9E+09,9E+09,9E+09,9E+09]];
    CONST robtarget Target_LetFron4_530:=[[-41.799,-124.084,66.777],[0.492892784,0.289203693,0.528592352,0.627700607],[0,0,0,0],[9E+09,9E+09,9E+09,9E+09,9E+09,9E+09]];
    CONST robtarget Target_LetFron4_540:=[[-51.881,-144.07,66.763],[0.492892784,0.289203693,0.528592352,0.627700607],[0,0,0,0],[9E+09,9E+09,9E+09,9E+09,9E+09,9E+09]];
    CONST robtarget Target_LetFron4_550:=[[-65.929,-140.725,71.706],[0.492892784,0.289203693,0.528592352,0.627700607],[0,0,0,0],[9E+09,9E+09,9E+09,9E+09,9E+09,9E+09]];
    CONST robtarget Target_LetFron4_560:=[[-55.929,-120.725,71.706],[0.492892784,0.289203693,0.528592352,0.627700607],[0,0,0,0],[9E+09,9E+09,9E+09,9E+09,9E+09,9E+09]];
    CONST robtarget Target_LetFron4_570:=[[-58.219,-120.014,72.135],[0.492892784,0.289203693,0.528592352,0.627700607],[0,0,0,0],[9E+09,9E+09,9E+09,9E+09,9E+09,9E+09]];
    CONST robtarget Target_LetFron4_580:=[[-59.351,-119.645,73.056],[0.492892784,0.289203693,0.528592352,0.627700607],[0,0,0,0],[9E+09,9E+09,9E+09,9E+09,9E+09,9E+09]];
    CONST robtarget Target_LetFron4_590:=[[-60.341,-119.312,74.807],[0.492892784,0.289203693,0.528592352,0.627700607],[0,0,0,0],[9E+09,9E+09,9E+09,9E+09,9E+09,9E+09]];
    CONST robtarget Target_LetFron4_600:=[[-60.436,-119.279,77.772],[0.492892784,0.289203693,0.528592352,0.627700607],[0,0,0,0],[9E+09,9E+09,9E+09,9E+09,9E+09,9E+09]];
    CONST robtarget Target_LetFron4_610:=[[-59.958,-119.441,79.76],[0.492892784,0.289203693,0.528592352,0.627700607],[0,0,0,0],[9E+09,9E+09,9E+09,9E+09,9E+09,9E+09]];
    CONST robtarget Target_LetFron4_620:=[[-59.173,-119.703,81.075],[0.492892784,0.289203693,0.528592352,0.627700607],[0,0,0,0],[9E+09,9E+09,9E+09,9E+09,9E+09,9E+09]];
    CONST robtarget Target_LetFron4_630:=[[-57.768,-120.156,81.941],[0.492892784,0.289203693,0.528592352,0.627700607],[0,0,0,0],[9E+09,9E+09,9E+09,9E+09,9E+09,9E+09]];
    CONST robtarget Target_LetFron4_640:=[[-55.396,-120.883,82.352],[0.492892784,0.289203693,0.528592352,0.627700607],[0,0,0,0],[9E+09,9E+09,9E+09,9E+09,9E+09,9E+09]];
    CONST robtarget Target_LetFron4_650:=[[-53.457,-121.439,81.782],[0.492892784,0.289203693,0.528592352,0.627700607],[0,0,0,0],[9E+09,9E+09,9E+09,9E+09,9E+09,9E+09]];
    CONST robtarget Target_LetFron4_660:=[[-52.512,-121.698,80.942],[0.492892784,0.289203693,0.528592352,0.627700607],[0,0,0,0],[9E+09,9E+09,9E+09,9E+09,9E+09,9E+09]];
    CONST robtarget Target_LetFron4_670:=[[-51.562,-121.95,79.035],[0.492892784,0.289203693,0.528592352,0.627700607],[0,0,0,0],[9E+09,9E+09,9E+09,9E+09,9E+09,9E+09]];
    CONST robtarget Target_LetFron4_680:=[[-51.38,-121.997,76.684],[0.492892784,0.289203693,0.528592352,0.627700607],[0,0,0,0],[9E+09,9E+09,9E+09,9E+09,9E+09,9E+09]];
    CONST robtarget Target_LetFron4_690:=[[-51.802,-121.887,74.523],[0.492892784,0.289203693,0.528592352,0.627700607],[0,0,0,0],[9E+09,9E+09,9E+09,9E+09,9E+09,9E+09]];
    CONST robtarget Target_LetFron4_700:=[[-52.915,-121.589,72.793],[0.492892784,0.289203693,0.528592352,0.627700607],[0,0,0,0],[9E+09,9E+09,9E+09,9E+09,9E+09,9E+09]];
    CONST robtarget Target_LetFron4_710:=[[-54.387,-121.177,71.924],[0.492892784,0.289203693,0.528592352,0.627700607],[0,0,0,0],[9E+09,9E+09,9E+09,9E+09,9E+09,9E+09]];
    CONST robtarget Target_LetFron4_720:=[[-56.264,-120.624,71.706],[0.492892784,0.289203693,0.528592352,0.627700607],[0,0,0,0],[9E+09,9E+09,9E+09,9E+09,9E+09,9E+09]];
    CONST robtarget Target_LetFron4_730:=[[-66.307,-140.611,71.706],[0.492892784,0.289203693,0.528592352,0.627700607],[0,0,0,0],[9E+09,9E+09,9E+09,9E+09,9E+09,9E+09]];
    CONST robtarget Target_LetFron4_740:=[[-77.909,-136.454,71.976],[0.492892784,0.289203693,0.528592352,0.627700607],[0,0,0,0],[9E+09,9E+09,9E+09,9E+09,9E+09,9E+09]];
    CONST robtarget Target_LetFron4_750:=[[-67.909,-116.454,71.976],[0.492892784,0.289203693,0.528592352,0.627700607],[0,0,0,0],[9E+09,9E+09,9E+09,9E+09,9E+09,9E+09]];
    CONST robtarget Target_LetFron4_760:=[[-61.598,-118.875,72.196],[0.492892784,0.289203693,0.528592352,0.627700607],[0,0,0,0],[9E+09,9E+09,9E+09,9E+09,9E+09,9E+09]];
    CONST robtarget Target_LetFron4_770:=[[-63.153,-118.315,71.808],[0.492892784,0.289203693,0.528592352,0.627700607],[0,0,0,0],[9E+09,9E+09,9E+09,9E+09,9E+09,9E+09]];
    CONST robtarget Target_LetFron4_780:=[[-63.249,-118.279,70.254],[0.492892784,0.289203693,0.528592352,0.627700607],[0,0,0,0],[9E+09,9E+09,9E+09,9E+09,9E+09,9E+09]];
    CONST robtarget Target_LetFron4_790:=[[-63.067,-118.347,80.357],[0.492892784,0.289203693,0.528592352,0.627700607],[0,0,0,0],[9E+09,9E+09,9E+09,9E+09,9E+09,9E+09]];
    CONST robtarget Target_LetFron4_800:=[[-63.524,-118.178,81.429],[0.492892784,0.289203693,0.528592352,0.627700607],[0,0,0,0],[9E+09,9E+09,9E+09,9E+09,9E+09,9E+09]];
    CONST robtarget Target_LetFron4_810:=[[-64.207,-117.922,81.987],[0.492892784,0.289203693,0.528592352,0.627700607],[0,0,0,0],[9E+09,9E+09,9E+09,9E+09,9E+09,9E+09]];
    CONST robtarget Target_LetFron4_820:=[[-65.492,-117.428,82.371],[0.492892784,0.289203693,0.528592352,0.627700607],[0,0,0,0],[9E+09,9E+09,9E+09,9E+09,9E+09,9E+09]];
    CONST robtarget Target_LetFron4_830:=[[-68.17,-116.346,81.741],[0.492892784,0.289203693,0.528592352,0.627700607],[0,0,0,0],[9E+09,9E+09,9E+09,9E+09,9E+09,9E+09]];
    CONST robtarget Target_LetFron4_840:=[[-78.17,-136.346,81.741],[0.492892784,0.289203693,0.528592352,0.627700607],[0,0,0,0],[9E+09,9E+09,9E+09,9E+09,9E+09,9E+09]];
    CONST robtarget Target_LetFron4_850:=[[-80.679,-135.265,82.097],[0.492892784,0.289203693,0.528592352,0.627700607],[0,0,0,0],[9E+09,9E+09,9E+09,9E+09,9E+09,9E+09]];
    CONST robtarget Target_LetFron4_860:=[[-70.679,-115.265,82.097],[0.492892784,0.289203693,0.528592352,0.627700607],[0,0,0,0],[9E+09,9E+09,9E+09,9E+09,9E+09,9E+09]];
    CONST robtarget Target_LetFron4_870:=[[-71.109,-115.074,71.804],[0.492892784,0.289203693,0.528592352,0.627700607],[0,0,0,0],[9E+09,9E+09,9E+09,9E+09,9E+09,9E+09]];
    CONST robtarget Target_LetFron4_880:=[[-81.109,-135.074,71.804],[0.492892784,0.289203693,0.528592352,0.627700607],[0,0,0,0],[9E+09,9E+09,9E+09,9E+09,9E+09,9E+09]];
    CONST robtarget Target_LetFron4_890:=[[-80.89,-135.172,67.298],[0.492892784,0.289203693,0.528592352,0.627700607],[0,0,0,0],[9E+09,9E+09,9E+09,9E+09,9E+09,9E+09]];
    CONST robtarget Target_LetFron4_900:=[[-70.89,-115.172,67.298],[0.492892784,0.289203693,0.528592352,0.627700607],[0,0,0,0],[9E+09,9E+09,9E+09,9E+09,9E+09,9E+09]];
    CONST robtarget Target_LetFron4_910:=[[-80.89,-135.172,67.298],[0.492892784,0.289203693,0.528592352,0.627700607],[0,0,0,0],[9E+09,9E+09,9E+09,9E+09,9E+09,9E+09]];
    CONST robtarget Target_LetFron4_920:=[[-83.841,-133.81,72.741],[0.492892784,0.289203693,0.528592352,0.627700607],[0,0,0,0],[9E+09,9E+09,9E+09,9E+09,9E+09,9E+09]];
    CONST robtarget Target_LetFron4_930:=[[-73.841,-113.81,72.741],[0.492892784,0.289203693,0.528592352,0.627700607],[0,0,0,0],[9E+09,9E+09,9E+09,9E+09,9E+09,9E+09]];
    CONST robtarget Target_LetFron4_940:=[[-80.391,-110.444,72.677],[0.492892784,0.289203693,0.528592352,0.627700607],[0,0,0,0],[9E+09,9E+09,9E+09,9E+09,9E+09,9E+09]];
    CONST robtarget Target_LetFron4_950:=[[-73.709,-113.873,81.484],[0.492892784,0.289203693,0.528592352,0.627700607],[0,0,0,0],[9E+09,9E+09,9E+09,9E+09,9E+09,9E+09]];
    CONST robtarget Target_LetFron4_960:=[[-80.618,-110.318,81.343],[0.492892784,0.289203693,0.528592352,0.627700607],[0,0,0,0],[9E+09,9E+09,9E+09,9E+09,9E+09,9E+09]];
    CONST robtarget Target_LetFron4_970:=[[-90.618,-130.318,81.343],[0.492892784,0.289203693,0.528592352,0.627700607],[0,0,0,0],[9E+09,9E+09,9E+09,9E+09,9E+09,9E+09]];
    CONST robtarget Target_LetFron4_980:=[[-96.912,-126.583,76.384],[0.492892784,0.289203693,0.528592352,0.627700607],[0,0,0,0],[9E+09,9E+09,9E+09,9E+09,9E+09,9E+09]];
    CONST robtarget Target_LetFron4_990:=[[-86.912,-106.583,76.384],[0.492892784,0.289203693,0.528592352,0.627700607],[0,0,0,0],[9E+09,9E+09,9E+09,9E+09,9E+09,9E+09]];
    CONST robtarget Target_LetFron4_1000:=[[-84.485,-108.082,76.613],[0.492892784,0.289203693,0.528592352,0.627700607],[0,0,0,0],[9E+09,9E+09,9E+09,9E+09,9E+09,9E+09]];
    CONST robtarget Target_LetFron4_1010:=[[-83.791,-108.494,77.082],[0.492892784,0.289203693,0.528592352,0.627700607],[0,0,0,0],[9E+09,9E+09,9E+09,9E+09,9E+09,9E+09]];
    CONST robtarget Target_LetFron4_1020:=[[-82.966,-108.983,77.537],[0.492892784,0.289203693,0.528592352,0.627700607],[0,0,0,0],[9E+09,9E+09,9E+09,9E+09,9E+09,9E+09]];
    CONST robtarget Target_LetFron4_1030:=[[-82.308,-109.365,78.42],[0.492892784,0.289203693,0.528592352,0.627700607],[0,0,0,0],[9E+09,9E+09,9E+09,9E+09,9E+09,9E+09]];
    CONST robtarget Target_LetFron4_1040:=[[-82.086,-109.491,80.116],[0.492892784,0.289203693,0.528592352,0.627700607],[0,0,0,0],[9E+09,9E+09,9E+09,9E+09,9E+09,9E+09]];
    CONST robtarget Target_LetFron4_1050:=[[-82.373,-109.326,81.085],[0.492892784,0.289203693,0.528592352,0.627700607],[0,0,0,0],[9E+09,9E+09,9E+09,9E+09,9E+09,9E+09]];
    CONST robtarget Target_LetFron4_1060:=[[-83.125,-108.889,81.922],[0.492892784,0.289203693,0.528592352,0.627700607],[0,0,0,0],[9E+09,9E+09,9E+09,9E+09,9E+09,9E+09]];
    CONST robtarget Target_LetFron4_1070:=[[-84.166,-108.273,82.32],[0.492892784,0.289203693,0.528592352,0.627700607],[0,0,0,0],[9E+09,9E+09,9E+09,9E+09,9E+09,9E+09]];
    CONST robtarget Target_LetFron4_1080:=[[-85.539,-107.441,82.127],[0.492892784,0.289203693,0.528592352,0.627700607],[0,0,0,0],[9E+09,9E+09,9E+09,9E+09,9E+09,9E+09]];
    CONST robtarget Target_LetFron4_1090:=[[-87.047,-106.497,81.2],[0.492892784,0.289203693,0.528592352,0.627700607],[0,0,0,0],[9E+09,9E+09,9E+09,9E+09,9E+09,9E+09]];
    CONST robtarget Target_LetFron4_1100:=[[-87.357,-106.3,82.283],[0.492892784,0.289203693,0.528592352,0.627700607],[0,0,0,0],[9E+09,9E+09,9E+09,9E+09,9E+09,9E+09]];
    CONST robtarget Target_LetFron4_1110:=[[-88.5,-105.56,82.045],[0.492892784,0.289203693,0.528592352,0.627700607],[0,0,0,0],[9E+09,9E+09,9E+09,9E+09,9E+09,9E+09]];
    CONST robtarget Target_LetFron4_1120:=[[-88.455,-105.589,74.61],[0.492892784,0.289203693,0.528592352,0.627700607],[0,0,0,0],[9E+09,9E+09,9E+09,9E+09,9E+09,9E+09]];
    CONST robtarget Target_LetFron4_1130:=[[-88.089,-105.827,73.106],[0.492892784,0.289203693,0.528592352,0.627700607],[0,0,0,0],[9E+09,9E+09,9E+09,9E+09,9E+09,9E+09]];
    CONST robtarget Target_LetFron4_1140:=[[-87.203,-106.397,72.116],[0.492892784,0.289203693,0.528592352,0.627700607],[0,0,0,0],[9E+09,9E+09,9E+09,9E+09,9E+09,9E+09]];
    CONST robtarget Target_LetFron4_1150:=[[-86.231,-107.012,71.706],[0.492892784,0.289203693,0.528592352,0.627700607],[0,0,0,0],[9E+09,9E+09,9E+09,9E+09,9E+09,9E+09]];
    CONST robtarget Target_LetFron4_1160:=[[-84.89,-107.838,71.741],[0.492892784,0.289203693,0.528592352,0.627700607],[0,0,0,0],[9E+09,9E+09,9E+09,9E+09,9E+09,9E+09]];
    CONST robtarget Target_LetFron4_1170:=[[-83.178,-108.859,72.224],[0.492892784,0.289203693,0.528592352,0.627700607],[0,0,0,0],[9E+09,9E+09,9E+09,9E+09,9E+09,9E+09]];
    CONST robtarget Target_LetFron4_1180:=[[-82.293,-109.373,72.583],[0.492892784,0.289203693,0.528592352,0.627700607],[0,0,0,0],[9E+09,9E+09,9E+09,9E+09,9E+09,9E+09]];
    CONST robtarget Target_LetFron4_1190:=[[-82.795,-109.082,73.885],[0.492892784,0.289203693,0.528592352,0.627700607],[0,0,0,0],[9E+09,9E+09,9E+09,9E+09,9E+09,9E+09]];
    CONST robtarget Target_LetFron4_1200:=[[-86.405,-106.902,73.751],[0.492892784,0.289203693,0.528592352,0.627700607],[0,0,0,0],[9E+09,9E+09,9E+09,9E+09,9E+09,9E+09]];
    CONST robtarget Target_LetFron4_1210:=[[-86.912,-106.583,76.365],[0.492892784,0.289203693,0.528592352,0.627700607],[0,0,0,0],[9E+09,9E+09,9E+09,9E+09,9E+09,9E+09]];
    CONST robtarget Target_LetFron4_1220:=[[-96.912,-126.583,76.365],[0.492892784,0.289203693,0.528592352,0.627700607],[0,0,0,0],[9E+09,9E+09,9E+09,9E+09,9E+09,9E+09]];
    CONST robtarget Target_LetFron4_1230:=[[-106.135,-120.138,71.999],[0.492892784,0.289203693,0.528592352,0.627700607],[0,0,0,0],[9E+09,9E+09,9E+09,9E+09,9E+09,9E+09]];
    CONST robtarget Target_LetFron4_1240:=[[-96.135,-100.138,72],[0.492892784,0.289203693,0.528592352,0.627700607],[0,0,0,0],[9E+09,9E+09,9E+09,9E+09,9E+09,9E+09]];
    CONST robtarget Target_LetFron4_1250:=[[-93.898,-101.817,71.706],[0.492892784,0.289203693,0.528592352,0.627700607],[0,0,0,0],[9E+09,9E+09,9E+09,9E+09,9E+09,9E+09]];
    CONST robtarget Target_LetFron4_1260:=[[-92.976,-102.487,72.044],[0.492892784,0.289203693,0.528592352,0.627700607],[0,0,0,0],[9E+09,9E+09,9E+09,9E+09,9E+09,9E+09]];
    CONST robtarget Target_LetFron4_1270:=[[-91.972,-103.201,72.746],[0.492892784,0.289203693,0.528592352,0.627700607],[0,0,0,0],[9E+09,9E+09,9E+09,9E+09,9E+09,9E+09]];
    CONST robtarget Target_LetFron4_1280:=[[-91.003,-103.877,74.083],[0.492892784,0.289203693,0.528592352,0.627700607],[0,0,0,0],[9E+09,9E+09,9E+09,9E+09,9E+09,9E+09]];
    CONST robtarget Target_LetFron4_1290:=[[-90.49,-104.229,75.778],[0.492892784,0.289203693,0.528592352,0.627700607],[0,0,0,0],[9E+09,9E+09,9E+09,9E+09,9E+09,9E+09]];
    CONST robtarget Target_LetFron4_1300:=[[-90.536,-104.197,78.92],[0.492892784,0.289203693,0.528592352,0.627700607],[0,0,0,0],[9E+09,9E+09,9E+09,9E+09,9E+09,9E+09]];
    CONST robtarget Target_LetFron4_1310:=[[-91.01,-103.872,80.48],[0.492892784,0.289203693,0.528592352,0.627700607],[0,0,0,0],[9E+09,9E+09,9E+09,9E+09,9E+09,9E+09]];
    CONST robtarget Target_LetFron4_1320:=[[-91.985,-103.192,81.757],[0.492892784,0.289203693,0.528592352,0.627700607],[0,0,0,0],[9E+09,9E+09,9E+09,9E+09,9E+09,9E+09]];
    CONST robtarget Target_LetFron4_1330:=[[-93.53,-102.086,82.389],[0.492892784,0.289203693,0.528592352,0.627700607],[0,0,0,0],[9E+09,9E+09,9E+09,9E+09,9E+09,9E+09]];
    CONST robtarget Target_LetFron4_1340:=[[-95.059,-100.955,82.014],[0.492892784,0.289203693,0.528592352,0.627700607],[0,0,0,0],[9E+09,9E+09,9E+09,9E+09,9E+09,9E+09]];
    CONST robtarget Target_LetFron4_1350:=[[-96.116,-100.153,81.394],[0.492892784,0.289203693,0.528592352,0.627700607],[0,0,0,0],[9E+09,9E+09,9E+09,9E+09,9E+09,9E+09]];
    CONST robtarget Target_LetFron4_1360:=[[-96.817,-99.61,82.324],[0.492892784,0.289203693,0.528592352,0.627700607],[0,0,0,0],[9E+09,9E+09,9E+09,9E+09,9E+09,9E+09]];
    CONST robtarget Target_LetFron4_1370:=[[-97.307,-99.227,82.179],[0.492892784,0.289203693,0.528592352,0.627700607],[0,0,0,0],[9E+09,9E+09,9E+09,9E+09,9E+09,9E+09]];
    CONST robtarget Target_LetFron4_1380:=[[-97.057,-99.423,66.726],[0.492892784,0.289203693,0.528592352,0.627700607],[0,0,0,0],[9E+09,9E+09,9E+09,9E+09,9E+09,9E+09]];
    CONST robtarget Target_LetFron4_1390:=[[-107.154,-119.348,66.706],[0.492892784,0.289203693,0.528592352,0.627700607],[0,0,0,0],[9E+09,9E+09,9E+09,9E+09,9E+09,9E+09]];
    CONST robtarget Target_LetFron4_1400:=[[-112.893,-114.561,71.706],[0.492892784,0.289203693,0.528592352,0.627700607],[0,0,0,0],[9E+09,9E+09,9E+09,9E+09,9E+09,9E+09]];
    CONST robtarget Target_LetFron4_1410:=[[-102.893,-94.561,71.706],[0.492892784,0.289203693,0.528592352,0.627700607],[0,0,0,0],[9E+09,9E+09,9E+09,9E+09,9E+09,9E+09]];
    CONST robtarget Target_LetFron4_1420:=[[-101.562,-95.724,72.214],[0.492892784,0.289203693,0.528592352,0.627700607],[0,0,0,0],[9E+09,9E+09,9E+09,9E+09,9E+09,9E+09]];
    CONST robtarget Target_LetFron4_1430:=[[-100.733,-96.432,72.868],[0.492892784,0.289203693,0.528592352,0.627700607],[0,0,0,0],[9E+09,9E+09,9E+09,9E+09,9E+09,9E+09]];
    CONST robtarget Target_LetFron4_1440:=[[-100.12,-96.947,73.973],[0.492892784,0.289203693,0.528592352,0.627700607],[0,0,0,0],[9E+09,9E+09,9E+09,9E+09,9E+09,9E+09]];
    CONST robtarget Target_LetFron4_1450:=[[-99.609,-97.371,75.571],[0.492892784,0.289203693,0.528592352,0.627700607],[0,0,0,0],[9E+09,9E+09,9E+09,9E+09,9E+09,9E+09]];
    CONST robtarget Target_LetFron4_1460:=[[-99.576,-97.398,77.889],[0.492892784,0.289203693,0.528592352,0.627700607],[0,0,0,0],[9E+09,9E+09,9E+09,9E+09,9E+09,9E+09]];
    CONST robtarget Target_LetFron4_1470:=[[-99.778,-97.232,79.518],[0.492892784,0.289203693,0.528592352,0.627700607],[0,0,0,0],[9E+09,9E+09,9E+09,9E+09,9E+09,9E+09]];
    CONST robtarget Target_LetFron4_1480:=[[-100.899,-96.29,81.443],[0.492892784,0.289203693,0.528592352,0.627700607],[0,0,0,0],[9E+09,9E+09,9E+09,9E+09,9E+09,9E+09]];
    CONST robtarget Target_LetFron4_1490:=[[-101.954,-95.385,82.187],[0.492892784,0.289203693,0.528592352,0.627700607],[0,0,0,0],[9E+09,9E+09,9E+09,9E+09,9E+09,9E+09]];
    CONST robtarget Target_LetFron4_1500:=[[-103.655,-93.881,82.389],[0.492892784,0.289203693,0.528592352,0.627700607],[0,0,0,0],[9E+09,9E+09,9E+09,9E+09,9E+09,9E+09]];
    CONST robtarget Target_LetFron4_1510:=[[-104.961,-92.688,81.737],[0.492892784,0.289203693,0.528592352,0.627700607],[0,0,0,0],[9E+09,9E+09,9E+09,9E+09,9E+09,9E+09]];
    CONST robtarget Target_LetFron4_1520:=[[-105.958,-91.753,80.398],[0.492892784,0.289203693,0.528592352,0.627700607],[0,0,0,0],[9E+09,9E+09,9E+09,9E+09,9E+09,9E+09]];
    CONST robtarget Target_LetFron4_1530:=[[-106.491,-91.246,79.13],[0.492892784,0.289203693,0.528592352,0.627700607],[0,0,0,0],[9E+09,9E+09,9E+09,9E+09,9E+09,9E+09]];
    CONST robtarget Target_LetFron4_1540:=[[-106.694,-91.051,77.754],[0.492892784,0.289203693,0.528592352,0.627700607],[0,0,0,0],[9E+09,9E+09,9E+09,9E+09,9E+09,9E+09]];
    CONST robtarget Target_LetFron4_1550:=[[-106.54,-91.198,75.105],[0.492892784,0.289203693,0.528592352,0.627700607],[0,0,0,0],[9E+09,9E+09,9E+09,9E+09,9E+09,9E+09]];
    CONST robtarget Target_LetFron4_1560:=[[-105.799,-91.904,73.056],[0.492892784,0.289203693,0.528592352,0.627700607],[0,0,0,0],[9E+09,9E+09,9E+09,9E+09,9E+09,9E+09]];
    CONST robtarget Target_LetFron4_1570:=[[-104.82,-92.818,72.044],[0.492892784,0.289203693,0.528592352,0.627700607],[0,0,0,0],[9E+09,9E+09,9E+09,9E+09,9E+09,9E+09]];
    CONST robtarget Target_LetFron4_1580:=[[-103.639,-93.895,71.706],[0.492892784,0.289203693,0.528592352,0.627700607],[0,0,0,0],[9E+09,9E+09,9E+09,9E+09,9E+09,9E+09]];
    CONST robtarget Target_LetFron4_1590:=[[-103.035,-94.436,71.706],[0.492892784,0.289203693,0.528592352,0.627700607],[0,0,0,0],[9E+09,9E+09,9E+09,9E+09,9E+09,9E+09]];
    CONST robtarget Target_LetFron4_1600:=[[-113.035,-114.436,71.706],[0.492892784,0.289203693,0.528592352,0.627700607],[0,0,0,0],[9E+09,9E+09,9E+09,9E+09,9E+09,9E+09]];
    CONST robtarget Target_LetFron4_1610:=[[-117.938,-109.837,81.072],[0.492892784,0.289203693,0.528592352,0.627700607],[0,0,0,0],[9E+09,9E+09,9E+09,9E+09,9E+09,9E+09]];
    CONST robtarget Target_LetFron4_1620:=[[-107.938,-89.837,81.072],[0.492892784,0.289203693,0.528592352,0.627700607],[0,0,0,0],[9E+09,9E+09,9E+09,9E+09,9E+09,9E+09]];
    CONST robtarget Target_LetFron4_1630:=[[-110.081,-87.662,82.389],[0.492892784,0.289203693,0.528592352,0.627700607],[0,0,0,0],[9E+09,9E+09,9E+09,9E+09,9E+09,9E+09]];
    CONST robtarget Target_LetFron4_1640:=[[-110.858,-86.848,82.288],[0.492892784,0.289203693,0.528592352,0.627700607],[0,0,0,0],[9E+09,9E+09,9E+09,9E+09,9E+09,9E+09]];
    CONST robtarget Target_LetFron4_1650:=[[-111.997,-85.626,81.57],[0.492892784,0.289203693,0.528592352,0.627700607],[0,0,0,0],[9E+09,9E+09,9E+09,9E+09,9E+09,9E+09]];
    CONST robtarget Target_LetFron4_1660:=[[-112.662,-84.897,80.511],[0.492892784,0.289203693,0.528592352,0.627700607],[0,0,0,0],[9E+09,9E+09,9E+09,9E+09,9E+09,9E+09]];
    CONST robtarget Target_LetFron4_1670:=[[-112.84,-84.7,79.426],[0.492892784,0.289203693,0.528592352,0.627700607],[0,0,0,0],[9E+09,9E+09,9E+09,9E+09,9E+09,9E+09]];
    CONST robtarget Target_LetFron4_1680:=[[-112.7,-84.856,78.197],[0.492892784,0.289203693,0.528592352,0.627700607],[0,0,0,0],[9E+09,9E+09,9E+09,9E+09,9E+09,9E+09]];
    CONST robtarget Target_LetFron4_1690:=[[-111.897,-85.734,76.939],[0.492892784,0.289203693,0.528592352,0.627700607],[0,0,0,0],[9E+09,9E+09,9E+09,9E+09,9E+09,9E+09]];
    CONST robtarget Target_LetFron4_1700:=[[-111.14,-86.548,76.411],[0.492892784,0.289203693,0.528592352,0.627700607],[0,0,0,0],[9E+09,9E+09,9E+09,9E+09,9E+09,9E+09]];
    CONST robtarget Target_LetFron4_1710:=[[-109.962,-87.786,75.717],[0.492892784,0.289203693,0.528592352,0.627700607],[0,0,0,0],[9E+09,9E+09,9E+09,9E+09,9E+09,9E+09]];
    CONST robtarget Target_LetFron4_1720:=[[-107.998,-89.777,74.886],[0.492892784,0.289203693,0.528592352,0.627700607],[0,0,0,0],[9E+09,9E+09,9E+09,9E+09,9E+09,9E+09]];
    CONST robtarget Target_LetFron4_1730:=[[-108.057,-89.718,73.869],[0.492892784,0.289203693,0.528592352,0.627700607],[0,0,0,0],[9E+09,9E+09,9E+09,9E+09,9E+09,9E+09]];
    CONST robtarget Target_LetFron4_1740:=[[-108.594,-89.183,72.718],[0.492892784,0.289203693,0.528592352,0.627700607],[0,0,0,0],[9E+09,9E+09,9E+09,9E+09,9E+09,9E+09]];
    CONST robtarget Target_LetFron4_1750:=[[-109.421,-88.344,72.026],[0.492892784,0.289203693,0.528592352,0.627700607],[0,0,0,0],[9E+09,9E+09,9E+09,9E+09,9E+09,9E+09]];
    CONST robtarget Target_LetFron4_1760:=[[-110.374,-87.356,71.732],[0.492892784,0.289203693,0.528592352,0.627700607],[0,0,0,0],[9E+09,9E+09,9E+09,9E+09,9E+09,9E+09]];
    CONST robtarget Target_LetFron4_1770:=[[-111.597,-86.059,71.794],[0.492892784,0.289203693,0.528592352,0.627700607],[0,0,0,0],[9E+09,9E+09,9E+09,9E+09,9E+09,9E+09]];
    CONST robtarget Target_LetFron4_1780:=[[-112.63,-84.933,72.718],[0.492892784,0.289203693,0.528592352,0.627700607],[0,0,0,0],[9E+09,9E+09,9E+09,9E+09,9E+09,9E+09]];
    CONST robtarget Target_LetFron4_1790:=[[-122.633,-104.929,72.696],[0.492892784,0.289203693,0.528592352,0.627700607],[0,0,0,0],[9E+09,9E+09,9E+09,9E+09,9E+09,9E+09]];
    CONST robtarget Target_LetFron4_1800:=[[-91.597,-85.059,-26.206],[0.443836724,0.190106418,0.616719914,0.621711396],[0,0,0,0],[9E+09,9E+09,9E+09,9E+09,9E+09,9E+09]];
    CONST robtarget Target_LetFron4_1810:=[[-92.63,-83.933,-25.282],[0.443836724,0.190106418,0.616719914,0.621711396],[0,0,0,0],[9E+09,9E+09,9E+09,9E+09,9E+09,9E+09]];
    CONST robtarget Target_LetFron4_1820:=[[-102.633,-103.929,-25.304],[0.443836724,0.190106418,0.616719914,0.621711396],[0,0,0,0],[9E+09,9E+09,9E+09,9E+09,9E+09,9E+09]];
    CONST robtarget p_contacto_labSIR{256}:=[Target_RobLab_20, Target_RobLab_30, Target_RobLab_40, Target_RobLab_50, Target_RobLab_60, Target_RobLab_70, Target_RobLab_80,
                                           Target_RobLab_90, Target_RobLab_100, Target_RobLab_110, Target_RobLab_120, Target_RobLab_130, Target_RobLab_140, Target_RobLab_150,
                                           Target_RobLab_160, Target_RobLab_170, Target_RobLab_180, Target_RobLab_190, Target_RobLab_200, Target_RobLab_210, Target_RobLab_220,
                                           Target_RobLab_230, Target_RobLab_240, Target_RobLab_250, Target_RobLab_260, Target_RobLab_280, Target_RobLab_290, Target_RobLab_300,
                                           Target_RobLab_310, Target_RobLab_320, Target_RobLab_330, Target_RobLab_340, Target_RobLab_350, Target_RobLab_360, Target_RobLab_370,
                                           Target_RobLab_380, Target_RobLab_390, Target_RobLab_400, Target_RobLab_410, Target_RobLab_420, Target_RobLab_430, Target_RobLab_440,
                                           Target_RobLab_450, Target_RobLab_460, Target_RobLab_470, Target_RobLab_480, Target_RobLab_490, Target_RobLab_500, Target_RobLab_510,
                                           Target_RobLab_520, Target_RobLab_530, Target_RobLab_540, Target_RobLab_550, Target_RobLab_560, Target_RobLab_570, Target_RobLab_580,
                                           Target_RobLab_590, Target_RobLab_600, Target_RobLab_610, Target_RobLab_620, Target_RobLab_630, Target_RobLab_640, Target_RobLab_650,
                                           Target_RobLab_660, Target_RobLab_670, Target_RobLab_680, Target_RobLab_690, Target_RobLab_700, Target_RobLab_710, Target_RobLab_720,
                                           Target_RobLab_730, Target_RobLab_740, Target_RobLab_750, Target_RobLab_760, Target_RobLab_770, Target_RobLab_780, Target_RobLab_790,
                                           Target_RobLab_800, Target_RobLab_810, Target_RobLab_820, Target_RobLab_830, Target_RobLab_840, Target_RobLab_850, Target_RobLab_860,
                                           Target_RobLab_870, Target_RobLab_880, Target_RobLab_890, Target_RobLab_900, Target_RobLab_910, Target_RobLab_920, Target_RobLab_930,
                                           Target_RobLab_940, Target_RobLab_950, Target_RobLab_960, Target_RobLab_980, Target_RobLab_990, Target_RobLab_1000, Target_RobLab_1010,
                                           Target_RobLab_1020, Target_RobLab_1030, Target_RobLab_1040, Target_RobLab_1050, Target_RobLab_1060, Target_RobLab_1070, Target_RobLab_1080,
                                           Target_RobLab_1090, Target_RobLab_1100, Target_RobLab_1110, Target_RobLab_1120, Target_RobLab_1130, Target_RobLab_1140, Target_RobLab_1160,
                                           Target_RobLab_1170, Target_RobLab_1180, Target_RobLab_1190, Target_RobLab_1200, Target_RobLab_1210, Target_RobLab_1220, Target_RobLab_1230,
                                           Target_RobLab_1240, Target_RobLab_1250, Target_RobLab_1260, Target_RobLab_1270, Target_RobLab_1280, Target_RobLab_1290, Target_RobLab_1310,
                                           Target_RobLab_1320, Target_RobLab_1330, Target_RobLab_1340, Target_RobLab_1350, Target_RobLab_1360, Target_RobLab_1380, Target_RobLab_1390,
                                           Target_RobLab_1400, Target_RobLab_1410, Target_RobLab_1420, Target_RobLab_1430, Target_RobLab_1450, Target_RobLab_1460, Target_RobLab_1470,
                                           Target_RobLab_1480, Target_RobLab_1490, Target_RobLab_1500, Target_RobLab_1520, Target_RobLab_1530, Target_RobLab_1540, Target_RobLab_1550,
                                           Target_RobLab_1560, Target_RobLab_1570, Target_RobLab_1590, Target_RobLab_1600, Target_RobLab_1610, Target_RobLab_1620, Target_RobLab_1630, Target_RobLab_1640,
                                           Target_RobLab_1660, Target_RobLab_1670, Target_RobLab_1680, Target_RobLab_1690, Target_RobLab_1700, Target_RobLab_1710, Target_Nom_L_20, Target_Nom_L_30,
                                           Target_Nom_L_40, Target_Nom_L_50, Target_Nom_L_60, Target_Nom_L_70, Target_Nom_L_80, Target_Nom_L_90, Target_Nom_L_100, Target_Nom_A_20, Target_Nom_A_30,
                                           Target_Nom_A_40, Target_Nom_A_50, Target_Nom_A_60, Target_Nom_A_70, Target_Nom_A_80, Target_Nom_A_90, Target_Nom_A_100, Target_Nom_A_110, Target_Nom_A_120,
                                           Target_Nom_A_130, Target_Nom_Aint_20, Target_Nom_Aint_30, Target_Nom_Aint_40, Target_Nom_Aint_50, Target_Nom_Aint_60, Target_Nom_Aint_70, Target_Nom_B_20,
                                           Target_Nom_B_30, Target_Nom_B_40, Target_Nom_B_50, Target_Nom_B_60, Target_Nom_B_70, Target_Nom_B_80, Target_Nom_B_90, Target_Nom_B_100, Target_Nom_B_110,
                                           Target_Nom_B_120, Target_Nom_Bint_20, Target_Nom_Bint_30, Target_Nom_Bint_40, Target_Nom_Bint_50, Target_Nom_Bint_60, Target_Nom_Bint_70, Target_Nom_R_20,
                                           Target_Nom_R_30, Target_Nom_R_40, Target_Nom_R_50, Target_Nom_R_60, Target_Nom_R_70, Target_Nom_R_80, Target_Nom_R_90, Target_Nom_R_100, Target_Nom_R_110,
                                           Target_Nom_R_120, Target_Nom_R_130, Target_Nom_R_140, Target_Nom_R_150, Target_Nom_Rint_20, Target_Nom_Rint_30, Target_Nom_Rint_40, Target_Nom_Rint_50,
                                           Target_Nom_Rint_60, Target_Nom_Rint_70, Target_Nom_Rint_80, Target_Nom_I_20, Target_Nom_I_30, Target_Nom_I_40, Target_Nom_I_50, Target_Nom_I_60, Target_Nom_I_70,
                                           Target_Nom_S_20, Target_Nom_S_30, Target_Nom_S_40, Target_Nom_S_50, Target_Nom_S_60, Target_Nom_S_70, Target_Nom_S_80, Target_Nom_S_90, Target_Nom_S_100, Target_Nom_S_110,
                                           Target_Nom_S_120, Target_Nom_S_130, Target_Nom_S_140, Target_Nom_S_150, Target_Nom_S_160, Target_Nom_S_170, Target_Nom_S_180, Target_Nom_S_190, Target_Nom_S_200, Target_Nom_S_210,
                                           Target_Nom_S_220, Target_Nom_S_230, Target_Nom_S_240, Target_Nom_S_250];
    CONST robtarget p_vacio_labSIR{19}:=[Target_RobLab_10, Target_RobLab_270, Target_RobLab_970, Target_RobLab_1150, Target_RobLab_1300, Target_RobLab_1370, Target_RobLab_1440,
                                        Target_RobLab_1510, Target_RobLab_1580, Target_RobLab_1650, Target_Nom_L_10, Target_Nom_A_10, Target_Nom_Aint_10, Target_Nom_B_10, Target_Nom_Bint_10,
                                        Target_Nom_R_10, Target_Nom_Rint_10, Target_Nom_I_10, Target_Nom_S_10];
    CONST robtarget p_contacto_labSIR_FrenteL{394}:=[Target_DibChip_20, Target_DibChip_30, Target_DibChip_40, Target_DibChip_50, Target_DibChip_60, Target_DibChip_70, Target_DibChip_80,
                                                     Target_DibChip_90, Target_DibChip_100, Target_DibChip_110, Target_DibChip_120, Target_DibChip_130, Target_DibChip_140, Target_DibChip_150,
                                                     Target_DibChip_160, Target_DibChip_170, Target_DibChip_180, Target_DibChip_190, Target_DibChip_200, Target_DibChip_210, Target_DibChip_220,
                                                     Target_DibChip_230, Target_DibChip_240, Target_DibChip_250, Target_DibChip_260, Target_DibChip_270, Target_DibChip_280, Target_DibChip_290,
                                                     Target_DibChip_300, Target_DibChip_310, Target_DibChip_320, Target_DibChip_330, Target_DibChip_340, Target_DibChip_350, Target_DibChip_360,
                                                     Target_DibChip_370, Target_DibChip_380, Target_DibChip_390, Target_DibChip_400, Target_DibChip_410, Target_DibChip_420, Target_DibChip_430,
                                                     Target_DibChip_440, Target_DibChip_450, Target_DibChip_460, Target_DibChip_470, Target_DibChip_480, Target_DibChip_490, Target_DibChip_500,
                                                     Target_DibChip_510, Target_DibChip_530, Target_DibChip_540, Target_DibChip_550, Target_DibChip_560, Target_DibChip_570, Target_DibChip_580,
                                                     Target_LetFron1_20, Target_LetFron1_30, Target_LetFron1_40, Target_LetFron1_50, Target_LetFron1_70, Target_LetFron1_80, Target_LetFron1_90,
                                                     Target_LetFron1_100, Target_LetFron1_110, Target_LetFron1_120, Target_LetFron1_130, Target_LetFron1_140, Target_LetFron1_150, Target_LetFron1_160,
                                                     Target_LetFron1_170, Target_LetFron1_180, Target_LetFron1_190, Target_LetFron1_200, Target_LetFron1_220, Target_LetFron1_230, Target_LetFron1_240,
                                                     Target_LetFron1_250, Target_LetFron1_260, Target_LetFron1_270, Target_LetFron1_280, Target_LetFron1_290, Target_LetFron1_300, Target_LetFron1_310,
                                                     Target_LetFron1_320, Target_LetFron1_330, Target_LetFron1_340, Target_LetFron1_350, Target_LetFron1_360, Target_LetFron1_370, Target_LetFron1_380,
                                                     Target_LetFron1_390, Target_LetFron1_410, Target_LetFron1_420, Target_LetFron1_430, Target_LetFron1_440, Target_LetFron1_450, Target_LetFron1_460,
                                                     Target_LetFron1_470, Target_LetFron1_480, Target_LetFron1_490, Target_LetFron1_500, Target_LetFron1_510, Target_LetFron1_520, Target_LetFron1_530,
                                                     Target_LetFron1_540, Target_LetFron1_550, Target_LetFron1_560, Target_LetFron1_570, Target_LetFron1_580, Target_LetFron1_590, Target_LetFron1_600,
                                                     Target_LetFron1_610, Target_LetFron1_620, Target_LetFron1_630, Target_LetFron1_640, Target_LetFron1_660, Target_LetFron1_670, Target_LetFron1_680,
                                                     Target_LetFron1_690, Target_LetFron1_700, Target_LetFron1_710, Target_LetFron1_730, Target_LetFron1_740, Target_LetFron1_750, Target_LetFron1_760,
                                                     Target_LetFron1_770, Target_LetFron1_780, Target_LetFron1_790, Target_LetFron1_800, Target_LetFron1_810, Target_LetFron1_820, Target_LetFron1_830,
                                                     Target_LetFron1_840, Target_LetFron1_850, Target_LetFron1_860, Target_LetFron1_870, Target_LetFron1_880, Target_LetFron1_890, Target_LetFron1_900,
                                                     Target_LetFron1_920, Target_LetFron1_930, Target_LetFron1_940, Target_LetFron1_950, Target_LetFron1_960, Target_LetFron1_970, Target_LetFron1_980,
                                                     Target_LetFron1_990, Target_LetFron1_1000, Target_LetFron1_1020, Target_LetFron1_1030, Target_LetFron1_1040, Target_LetFron1_1050, Target_LetFron1_1060,
                                                     Target_LetFron1_1070, Target_LetFron1_1080, Target_LetFron1_1090, Target_LetFron1_1100, Target_LetFron1_1110, Target_LetFron1_1120, Target_LetFron1_1130,
                                                     Target_LetFron1_1140, Target_LetFron1_1150, Target_LetFron1_1160, Target_LetFron1_1170, Target_LetFron1_1180, Target_LetFron1_1190, Target_LetFron1_1200,
                                                     Target_LetFron1_1210, Target_LetFron1_1220, Target_LetFron1_1230, Target_LetFron1_1240, Target_LetFron1_1250, Target_LetFron1_1260, Target_LetFron1_1280,
                                                     Target_LetFron1_1290, Target_LetFron1_1300, Target_LetFron1_1310, Target_LetFron1_1320, Target_LetFron1_1330, Target_LetFron1_1340, Target_LetFron1_1350,
                                                     Target_LetFron1_1360, Target_LetFron1_1380, Target_LetFron1_1390, Target_LetFron1_1400, Target_LetFron1_1420, Target_LetFron1_1430, Target_LetFron1_1450,
                                                     Target_LetFron1_1460, Target_LetFron1_1470, Target_LetFron1_1480, Target_LetFron1_1490, Target_LetFron1_1500, Target_LetFron1_1510, Target_LetFron1_1520,
                                                     Target_LetFron1_1530, Target_LetFron1_1540, Target_LetFron1_1550, Target_LetFron1_1560, Target_LetFron1_1570, Target_LetFron1_1580, Target_LetFron1_1590,
                                                     Target_LetFron1_1600, Target_LetFron1_1610, Target_LetFron1_1620, Target_LetFron1_1630, Target_LetFron1_1640, Target_LetFron1_1650, Target_LetFron1_1660,
                                                     Target_LetFron1_1670, Target_LetFron1_1680, Target_LetFron2_20, Target_LetFron2_30, Target_LetFron2_40, Target_LetFron2_50, Target_LetFron2_60,
                                                     Target_LetFron2_70, Target_LetFron2_80, Target_LetFron2_90, Target_LetFron2_100, Target_LetFron2_110, Target_LetFron2_120, Target_LetFron2_160,
                                                     Target_LetFron2_200, Target_LetFron2_210, Target_LetFron2_220, Target_LetFron2_230, Target_LetFron2_250, Target_LetFron2_260, Target_LetFron2_270,
                                                     Target_LetFron2_280, Target_LetFron2_290, Target_LetFron2_300, Target_LetFron2_310, Target_LetFron2_320, Target_LetFron2_330, Target_LetFron2_340,
                                                     Target_LetFron2_360, Target_LetFron2_370, Target_LetFron2_380, Target_LetFron2_390, Target_LetFron2_400, Target_LetFron2_410, Target_LetFron2_420,
                                                     Target_LetFron2_430, Target_LetFron2_440, Target_LetFron2_450, Target_LetFron2_460, Target_LetFron2_470, Target_LetFron2_480, Target_LetFron2_490,
                                                     Target_LetFron2_500, Target_LetFron2_510, Target_LetFron2_520, Target_LetFron2_530, Target_LetFron2_540, Target_LetFron2_550, Target_LetFron2_560,
                                                     Target_LetFron2_570, Target_LetFron2_580, Target_LetFron2_590, Target_LetFron2_610, Target_LetFron2_620, Target_LetFron2_630, Target_LetFron2_640,
                                                     Target_LetFron2_650, Target_LetFron2_660, Target_LetFron2_670, Target_LetFron2_680, Target_LetFron2_690, Target_LetFron2_700, Target_LetFron2_710,
                                                     Target_LetFron2_730, Target_LetFron2_740, Target_LetFron2_750, Target_LetFron2_760, Target_LetFron2_770, Target_LetFron2_780, Target_LetFron2_790,
                                                     Target_LetFron2_800, Target_LetFron2_810, Target_LetFron2_820, Target_LetFron2_830, Target_LetFron2_840, Target_LetFron2_850, Target_LetFron2_860,
                                                     Target_LetFron2_880, Target_LetFron2_890, Target_LetFron2_900, Target_LetFron2_910, Target_LetFron2_920, Target_LetFron2_940, Target_LetFron2_950,
                                                     Target_LetFron2_960, Target_LetFron2_970, Target_LetFron2_980, Target_LetFron2_990, Target_LetFron2_1000, Target_LetFron2_1010, Target_LetFron2_1020,
                                                     Target_LetFron2_1030, Target_LetFron2_1040, Target_LetFron2_1050, Target_LetFron2_1060, Target_LetFron2_1070, Target_LetFron2_1080, Target_LetFron2_1100,
                                                     Target_LetFron2_1110, Target_LetFron2_1120, Target_LetFron2_1130, Target_LetFron2_1140, Target_LetFron2_1150, Target_LetFron2_1160, Target_LetFron2_1170,
                                                     Target_LetFron2_1180, Target_LetFron2_1190, Target_LetFron2_1200, Target_LetFron2_1210, Target_LetFron2_1220, Target_LetFron2_1230, Target_LetFron2_1240,
                                                     Target_LetFron2_1250, Target_LetFron2_1260, Target_LetFron2_1270, Target_LetFron2_1280, Target_LetFron2_1290, Target_LetFron2_1300, Target_LetFron2_1310,
                                                     Target_LetFron2_1320, Target_LetFron2_1330, Target_LetFron2_1340, Target_LetFron2_1350, Target_LetFron2_1360, Target_LetFron2_1370, Target_LetFron2_1380,
                                                     Target_LetFron2_1390, Target_LetFron2_1400, Target_LetFron2_1410, Target_LetFron2_1420, Target_LetFron2_1430, Target_LetFron2_1450, Target_LetFron2_1460,
                                                     Target_LetFron2_1470, Target_LetFron2_1490, Target_LetFron2_1500, Target_LetFron2_1520, Target_LetFron2_1530, Target_LetFron2_1540, Target_LetFron2_1550,
                                                     Target_LetFron2_1570, Target_LetFron2_1580, Target_LetFron2_1590, Target_LetFron2_1600, Target_LetFron2_1610, Target_LetFron2_1620, Target_LetFron2_1630,
                                                     Target_LetFron2_1640, Target_LetFron2_1650, Target_LetFron2_1660, Target_LetFron2_1670, Target_LetFron2_1680, Target_LetFron2_1690, Target_LetFron2_1700,
                                                     Target_LetFron2_1710, Target_LetFron2_1720, Target_LetFron2_1730, Target_LetFron2_1740, Target_LetFron2_1750, Target_LetFron2_1760, Target_LetFron2_1780,
                                                     Target_LetFron2_1790, Target_LetFron2_1800, Target_LetFron2_1810, Target_LetFron2_1820, Target_LetFron2_1830, Target_LetFron2_1840, Target_LetFron2_1850,
                                                     Target_LetFron2_1860, Target_LetFron2_1880, Target_LetFron2_1890, Target_LetFron2_1900, Target_LetFron2_1910, Target_LetFron2_1920, Target_LetFron2_1930,
                                                     Target_LetFron2_1940, Target_LetFron2_1950, Target_LetFron2_1960, Target_LetFron2_1970, Target_LetFron2_1980, Target_LetFron2_1990, Target_LetFron2_2010,
                                                     Target_LetFron2_2020, Target_LetFron2_2030];
    CONST robtarget p_vacio_labSIR_FrenteL{27}:=[Target_DibChip_10, Target_DibChip_520, Target_LetFron1_10, Target_LetFron1_60, Target_LetFron1_210, Target_LetFron1_400, Target_LetFron1_650, Target_LetFron1_720,
                                                 Target_LetFron1_910, Target_LetFron1_1010, Target_LetFron1_1270, Target_LetFron1_1370, Target_LetFron1_1410, Target_LetFron1_1440, Target_LetFron2_10, Target_LetFron2_350,
                                                 Target_LetFron2_600, Target_LetFron2_720, Target_LetFron2_870, Target_LetFron2_1090, Target_LetFron2_1440, Target_LetFron2_1480, Target_LetFron2_1510, Target_LetFron2_1560,
                                                 Target_LetFron2_1770, Target_LetFron2_1870, Target_LetFron2_2000];
    CONST robtarget p_contacto_labSIR_FrenteR{448}:=[Target_DibEng_20, Target_DibEng_30, Target_DibEng_40, Target_DibEng_50, Target_DibEng_60, Target_DibEng_70, Target_DibEng_80, Target_DibEng_90, Target_DibEng_100,
                                                   Target_DibEng_110, Target_DibEng_120, Target_DibEng_130, Target_DibEng_140, Target_DibEng_150, Target_DibEng_160, Target_DibEng_170, Target_DibEng_180, Target_DibEng_190,
                                                   Target_DibEng_200, Target_DibEng_210, Target_DibEng_220, Target_DibEng_230, Target_DibEng_240, Target_DibEng_250, Target_DibEng_260, Target_DibEng_270, Target_DibEng_280,
                                                   Target_DibEng_290, Target_DibEng_300, Target_DibEng_310, Target_DibEng_320, Target_DibEng_330, Target_DibEng_340, Target_DibEng_350, Target_DibEng_360, Target_DibEng_370,
                                                   Target_DibEng_380, Target_DibEng_390, Target_DibEng_400, Target_DibEng_410, Target_DibEng_420, Target_DibEng_430, Target_DibEng_440, Target_DibEng_450, Target_DibEng_460,
                                                   Target_DibEng_470, Target_DibEng_480, Target_DibEng_490, Target_DibEng_500, Target_DibEng_510, Target_DibEng_520, Target_DibEng_530, Target_DibEng_540, Target_DibEng_550,
                                                   Target_DibEng_560, Target_DibEng_570, Target_DibEng_580, Target_DibEng_590, Target_DibEng_600, Target_DibEng_610, Target_DibEng_620, Target_DibEng_630, Target_DibEng_640,
                                                   Target_DibEng_650, Target_DibEng_660, Target_DibEng_670, Target_DibEng_680, Target_DibEng_690, Target_DibEng_700, Target_DibEng_710, Target_DibEng_720, Target_DibEng_730,
                                                   Target_DibEng_740, Target_DibEng_750, Target_DibEng_760, Target_DibEng_770, Target_DibEng_780, Target_DibEng_790, Target_DibEng_810, Target_DibEng_820, Target_DibEng_830,
                                                   Target_DibEng_840, Target_DibEng_850, Target_DibEng_860, Target_DibEng_870, Target_DibEng_880, Target_DibEng_890, Target_DibEng_900, Target_DibEng_910, Target_DibEng_920,
                                                   Target_DibEng_930, Target_DibEng_940, Target_DibEng_950, Target_DibEng_960, Target_DibEng_970, Target_DibEng_980, Target_DibEng_990, Target_LetFron3_20, Target_LetFron3_30,
                                                   Target_LetFron3_40, Target_LetFron3_50, Target_LetFron3_60, Target_LetFron3_70, Target_LetFron3_80, Target_LetFron3_90, Target_LetFron3_100, Target_LetFron3_110, Target_LetFron3_120,
                                                   Target_LetFron3_130, Target_LetFron3_140, Target_LetFron3_150, Target_LetFron3_160, Target_LetFron3_170, Target_LetFron3_180, Target_LetFron3_190, Target_LetFron3_200, Target_LetFron3_210,
                                                   Target_LetFron3_220, Target_LetFron3_230, Target_LetFron3_240, Target_LetFron3_250, Target_LetFron3_270, Target_LetFron3_280, Target_LetFron3_290, Target_LetFron3_300, Target_LetFron3_310,
                                                   Target_LetFron3_320, Target_LetFron3_330, Target_LetFron3_340, Target_LetFron3_350, Target_LetFron3_360, Target_LetFron3_370, Target_LetFron3_380, Target_LetFron3_390, Target_LetFron3_400,
                                                   Target_LetFron3_410, Target_LetFron3_420, Target_LetFron3_430, Target_LetFron3_440, Target_LetFron3_450, Target_LetFron3_460, Target_LetFron3_470, Target_LetFron3_480, Target_LetFron3_490,
                                                   Target_LetFron3_500, Target_LetFron3_510, Target_LetFron3_520, Target_LetFron3_530, Target_LetFron3_540, Target_LetFron3_550, Target_LetFron3_570, Target_LetFron3_580, Target_LetFron3_590,
                                                   Target_LetFron3_600, Target_LetFron3_610, Target_LetFron3_620, Target_LetFron3_630, Target_LetFron3_640, Target_LetFron3_650, Target_LetFron3_660, Target_LetFron3_670, Target_LetFron3_680,
                                                   Target_LetFron3_690, Target_LetFron3_710, Target_LetFron3_720, Target_LetFron3_730, Target_LetFron3_740, Target_LetFron3_750, Target_LetFron3_760, Target_LetFron3_770, Target_LetFron3_780,
                                                   Target_LetFron3_790, Target_LetFron3_800, Target_LetFron3_810, Target_LetFron3_820, Target_LetFron3_830, Target_LetFron3_840, Target_LetFron3_850, Target_LetFron3_860, Target_LetFron3_870,
                                                   Target_LetFron3_880, Target_LetFron3_890, Target_LetFron3_900, Target_LetFron3_910, Target_LetFron3_920, Target_LetFron3_930, Target_LetFron3_940, Target_LetFron3_960, Target_LetFron3_970,
                                                   Target_LetFron3_980, Target_LetFron3_990, Target_LetFron3_1000, Target_LetFron3_1010, Target_LetFron3_1020, Target_LetFron3_1030, Target_LetFron3_1040, Target_LetFron3_1050, Target_LetFron3_1060,
                                                   Target_LetFron3_1080, Target_LetFron3_1090, Target_LetFron3_1100, Target_LetFron3_1110, Target_LetFron3_1120, Target_LetFron3_1130, Target_LetFron3_1140, Target_LetFron3_1150, Target_LetFron3_1160,
                                                   Target_LetFron3_1170, Target_LetFron3_1180, Target_LetFron3_1190, Target_LetFron3_1200, Target_LetFron3_1210, Target_LetFron3_1220, Target_LetFron3_1230, Target_LetFron3_1240, Target_LetFron3_1250,
                                                   Target_LetFron3_1260, Target_LetFron3_1270, Target_LetFron3_1290, Target_LetFron3_1300, Target_LetFron3_1310, Target_LetFron3_1330, Target_LetFron3_1340, Target_LetFron3_1360, Target_LetFron3_1370,
                                                   Target_LetFron3_1380, Target_LetFron3_1390, Target_LetFron3_1400, Target_LetFron3_1410, Target_LetFron3_1420, Target_LetFron3_1430, Target_LetFron3_1440, Target_LetFron3_1450, Target_LetFron3_1460,
                                                   Target_LetFron3_1470, Target_LetFron3_1480, Target_LetFron3_1490, Target_LetFron3_1500, Target_LetFron3_1510, Target_LetFron3_1520, Target_LetFron3_1530, Target_LetFron3_1540, Target_LetFron3_1560,
                                                   Target_LetFron3_1570, Target_LetFron3_1580, Target_LetFron3_1590, Target_LetFron3_1600, Target_LetFron3_1610, Target_LetFron3_1620, Target_LetFron3_1630, Target_LetFron3_1640, Target_LetFron3_1650,
                                                   Target_LetFron3_1660, Target_LetFron3_1670, Target_LetFron3_1680, Target_LetFron3_1690, Target_LetFron3_1700, Target_LetFron3_1710, Target_LetFron3_1720, Target_LetFron3_1730, Target_LetFron3_1740,
                                                   Target_LetFron3_1750, Target_LetFron3_1760, Target_LetFron3_1770, Target_LetFron3_1790, Target_LetFron3_1800, Target_LetFron3_1810, Target_LetFron3_1820, Target_LetFron3_1830, Target_LetFron3_1840,
                                                   Target_LetFron3_1850, Target_LetFron3_1860, Target_LetFron3_1870, Target_LetFron3_1880, Target_LetFron3_1890, Target_LetFron3_1900, Target_LetFron3_1910, Target_LetFron3_1920, Target_LetFron3_1930,
                                                   Target_LetFron3_1940, Target_LetFron3_1950, Target_LetFron4_20, Target_LetFron4_30, Target_LetFron4_40, Target_LetFron4_50, Target_LetFron4_60, Target_LetFron4_70, Target_LetFron4_80, Target_LetFron4_90,
                                                   Target_LetFron4_100, Target_LetFron4_110, Target_LetFron4_120, Target_LetFron4_130, Target_LetFron4_150, Target_LetFron4_160, Target_LetFron4_170, Target_LetFron4_180, Target_LetFron4_190, Target_LetFron4_200,
                                                   Target_LetFron4_210, Target_LetFron4_220, Target_LetFron4_230, Target_LetFron4_240, Target_LetFron4_250, Target_LetFron4_260, Target_LetFron4_270, Target_LetFron4_280, Target_LetFron4_290, Target_LetFron4_300,
                                                   Target_LetFron4_310, Target_LetFron4_320, Target_LetFron4_330, Target_LetFron4_340, Target_LetFron4_350, Target_LetFron4_360, Target_LetFron4_370, Target_LetFron4_380, Target_LetFron4_400, Target_LetFron4_410,
                                                   Target_LetFron4_420, Target_LetFron4_430, Target_LetFron4_440, Target_LetFron4_450, Target_LetFron4_460, Target_LetFron4_470, Target_LetFron4_480, Target_LetFron4_490, Target_LetFron4_500, Target_LetFron4_510,
                                                   Target_LetFron4_520, Target_LetFron4_530, Target_LetFron4_540, Target_LetFron4_560, Target_LetFron4_570, Target_LetFron4_580, Target_LetFron4_590, Target_LetFron4_600, Target_LetFron4_610, Target_LetFron4_620,
                                                   Target_LetFron4_630, Target_LetFron4_640, Target_LetFron4_650, Target_LetFron4_660, Target_LetFron4_670, Target_LetFron4_680, Target_LetFron4_690, Target_LetFron4_700, Target_LetFron4_710, Target_LetFron4_720,
                                                   Target_LetFron4_730, Target_LetFron4_750, Target_LetFron4_760, Target_LetFron4_770, Target_LetFron4_780, Target_LetFron4_790, Target_LetFron4_800, Target_LetFron4_810, Target_LetFron4_820, Target_LetFron4_830,
                                                   Target_LetFron4_840, Target_LetFron4_860, Target_LetFron4_870, Target_LetFron4_880, Target_LetFron4_900, Target_LetFron4_910, Target_LetFron4_930, Target_LetFron4_940, Target_LetFron4_950, Target_LetFron4_960,
                                                   Target_LetFron4_970, Target_LetFron4_990, Target_LetFron4_1000, Target_LetFron4_1010, Target_LetFron4_1020, Target_LetFron4_1030, Target_LetFron4_1040, Target_LetFron4_1050, Target_LetFron4_1060, Target_LetFron4_1070,
                                                   Target_LetFron4_1080, Target_LetFron4_1090, Target_LetFron4_1100, Target_LetFron4_1110, Target_LetFron4_1120, Target_LetFron4_1130, Target_LetFron4_1140, Target_LetFron4_1150, Target_LetFron4_1160, Target_LetFron4_1170,
                                                   Target_LetFron4_1180, Target_LetFron4_1190, Target_LetFron4_1200, Target_LetFron4_1210, Target_LetFron4_1220, Target_LetFron4_1240, Target_LetFron4_1250, Target_LetFron4_1260, Target_LetFron4_1270, Target_LetFron4_1280,
                                                   Target_LetFron4_1290, Target_LetFron4_1300, Target_LetFron4_1310, Target_LetFron4_1320, Target_LetFron4_1330, Target_LetFron4_1340, Target_LetFron4_1350, Target_LetFron4_1360, Target_LetFron4_1370, Target_LetFron4_1380,
                                                   Target_LetFron4_1390, Target_LetFron4_1410, Target_LetFron4_1420, Target_LetFron4_1430, Target_LetFron4_1440, Target_LetFron4_1450, Target_LetFron4_1460, Target_LetFron4_1470, Target_LetFron4_1480, Target_LetFron4_1490,
                                                   Target_LetFron4_1500, Target_LetFron4_1510, Target_LetFron4_1520, Target_LetFron4_1530, Target_LetFron4_1540, Target_LetFron4_1550, Target_LetFron4_1560, Target_LetFron4_1570, Target_LetFron4_1580, Target_LetFron4_1590,
                                                   Target_LetFron4_1600, Target_LetFron4_1620, Target_LetFron4_1630, Target_LetFron4_1640, Target_LetFron4_1650, Target_LetFron4_1660, Target_LetFron4_1670, Target_LetFron4_1680, Target_LetFron4_1690, Target_LetFron4_1700,
                                                   Target_LetFron4_1710, Target_LetFron4_1720, Target_LetFron4_1730, Target_LetFron4_1740, Target_LetFron4_1750, Target_LetFron4_1760, Target_LetFron4_1770, Target_LetFron4_1780, Target_LetFron4_1790];
    CONST robtarget p_vacio_labSIR_FrenteR{25}:=[Target_DibEng_10, Target_DibEng_800, Target_LetFron3_10, Target_LetFron3_260, Target_LetFron3_560, Target_LetFron3_700, Target_LetFron3_950, Target_LetFron3_1070, Target_LetFron3_1280,
                                                Target_LetFron3_1320, Target_LetFron3_1350, Target_LetFron3_1550, Target_LetFron3_1780, Target_LetFron4_10, Target_LetFron4_140, Target_LetFron4_390, Target_LetFron4_550, Target_LetFron4_740,
                                                Target_LetFron4_850, Target_LetFron4_890, Target_LetFron4_920, Target_LetFron4_980, Target_LetFron4_1230, Target_LetFron4_1400, Target_LetFron4_1610];
    !PERS wobjdata WO_Pastel
    PROC Decorar_LABSIR(PERS wobjdata WO_Pastel)
        ReiniciarIndices;
        Path_Tapa_LabSIR WO_Pastel;
        Path_Frente_LabSIR WO_Pastel;
    ENDPROC

